PROGRAM prg_Piston
VAR
	fbPiston: FB_Piston;
	stPiston: ST_Piston;

	bPis_Next_P: BOOL;
	bPis_Next_N: BOOL;

	

	
	TON_0: TON;
	TON_1: TON;
	TON_2: TON;
	TON_3: TON;
	TON_4: TON;
	TON_5: TON;	
	i: INT;
END_VAR

act_InterLock();
act_Call_list_TanksMarinade();
act_Call_list_TanksColor();
act_Call_list_TanksCoolant();
act_Call_List_LineSource();
act_Call_List_LineTarget();
act_Call_list_CIP_SourceNTarget();
act_Call_list_CIP_Client();
act_Call_list_CIP_Tanks();
act_Call_list_Water();
act_Call_list_TriBlender_Selector();


IF bPis_Next_P THEN;
	m_Get_Next_P(iSel:=iPis_sel);
	bPis_Next_P:=FALSE;
END_IF

IF bPis_Next_N THEN;
	m_Get_Next_N(iSel:=iPis_sel);
	bPis_Next_N:=FALSE;
END_IF

FOR i:=0 TO E_Pis_Name.last DO
	ePisNameList:=i;
	arPisNameList[i]:=TO_STRING(ePisNameList);
END_FOR

ACTION act_Call_list_CIP_Client:
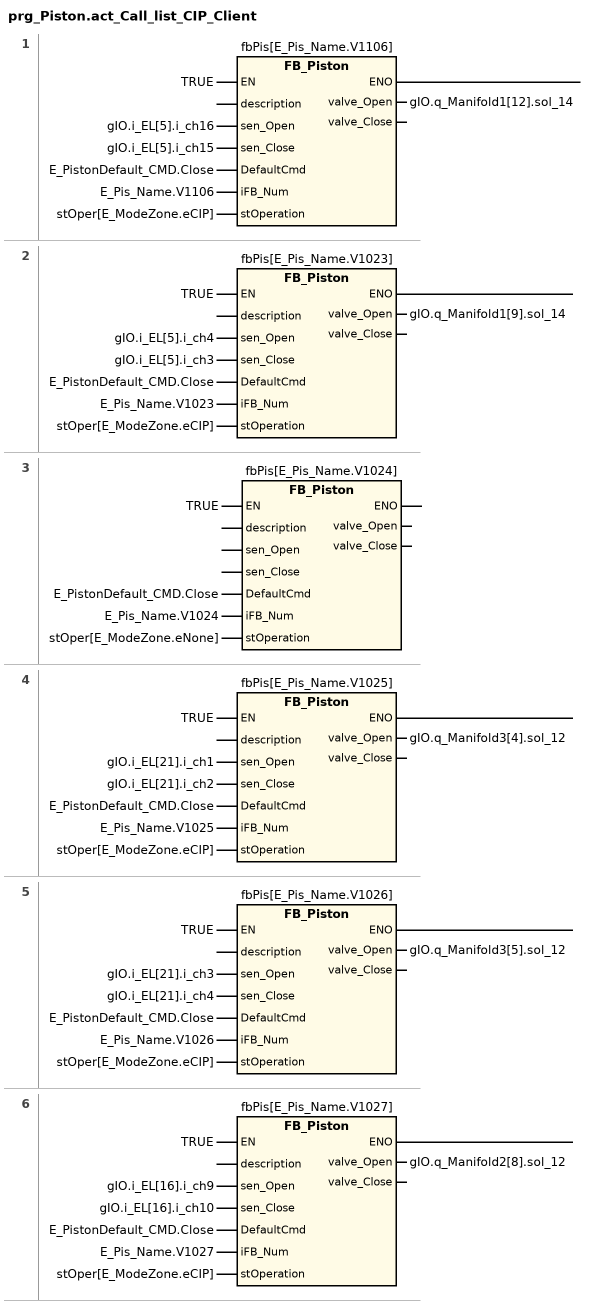
// NETWORK 1
fbPis[E_Pis_Name.V1106](
    sen_Open := gIO.i_EL[5].i_ch16,
    sen_Close := gIO.i_EL[5].i_ch15,
    DefaultCmd := E_PistonDefault_CMD.Close,
    iFB_Num := E_Pis_Name.V1106,
    stOperation := stOper[E_ModeZone.eCIP],
    valve_Open => gIO.q_Manifold1[12].sol_14); // FB_Piston

// NETWORK 2
fbPis[E_Pis_Name.V1023](
    sen_Open := gIO.i_EL[5].i_ch4,
    sen_Close := gIO.i_EL[5].i_ch3,
    DefaultCmd := E_PistonDefault_CMD.Close,
    iFB_Num := E_Pis_Name.V1023,
    stOperation := stOper[E_ModeZone.eCIP],
    valve_Open => gIO.q_Manifold1[9].sol_14); // FB_Piston

// NETWORK 3
fbPis[E_Pis_Name.V1024](
    DefaultCmd := E_PistonDefault_CMD.Close,
    iFB_Num := E_Pis_Name.V1024,
    stOperation := stOper[E_ModeZone.eNone]); // FB_Piston

// NETWORK 4
fbPis[E_Pis_Name.V1025](
    sen_Open := gIO.i_EL[21].i_ch1,
    sen_Close := gIO.i_EL[21].i_ch2,
    DefaultCmd := E_PistonDefault_CMD.Close,
    iFB_Num := E_Pis_Name.V1025,
    stOperation := stOper[E_ModeZone.eCIP],
    valve_Open => gIO.q_Manifold3[4].sol_12); // FB_Piston

// NETWORK 5
fbPis[E_Pis_Name.V1026](
    sen_Open := gIO.i_EL[21].i_ch3,
    sen_Close := gIO.i_EL[21].i_ch4,
    DefaultCmd := E_PistonDefault_CMD.Close,
    iFB_Num := E_Pis_Name.V1026,
    stOperation := stOper[E_ModeZone.eCIP],
    valve_Open => gIO.q_Manifold3[5].sol_12); // FB_Piston

// NETWORK 6
fbPis[E_Pis_Name.V1027](
    sen_Open := gIO.i_EL[16].i_ch9,
    sen_Close := gIO.i_EL[16].i_ch10,
    DefaultCmd := E_PistonDefault_CMD.Close,
    iFB_Num := E_Pis_Name.V1027,
    stOperation := stOper[E_ModeZone.eCIP],
    valve_Open => gIO.q_Manifold2[8].sol_12); // FB_Piston

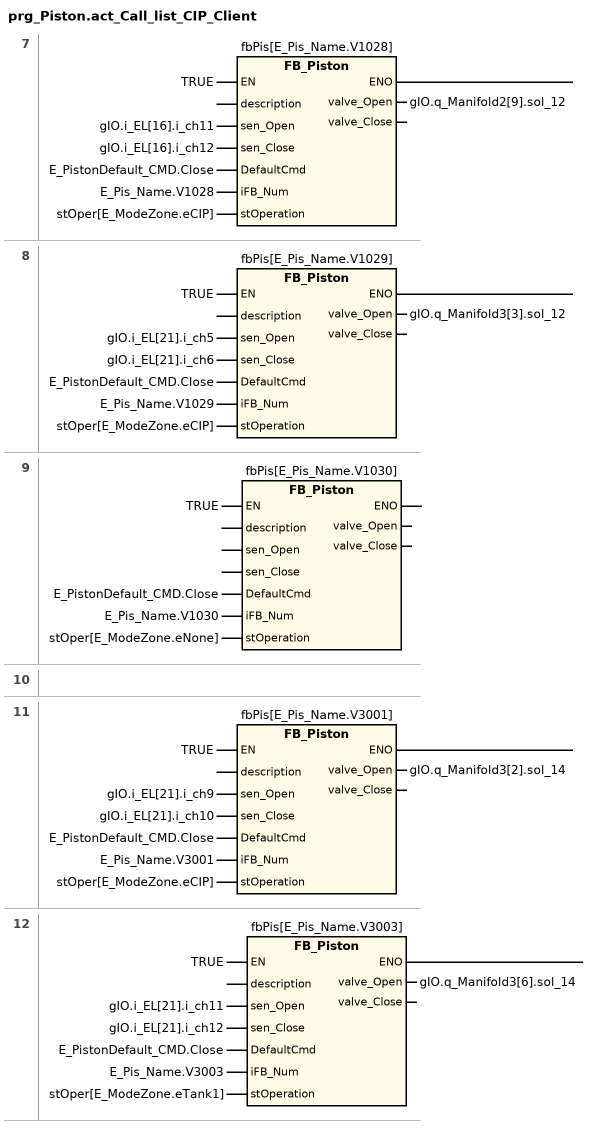
// NETWORK 7
fbPis[E_Pis_Name.V1028](
    sen_Open := gIO.i_EL[16].i_ch11,
    sen_Close := gIO.i_EL[16].i_ch12,
    DefaultCmd := E_PistonDefault_CMD.Close,
    iFB_Num := E_Pis_Name.V1028,
    stOperation := stOper[E_ModeZone.eCIP],
    valve_Open => gIO.q_Manifold2[9].sol_12); // FB_Piston

// NETWORK 8
fbPis[E_Pis_Name.V1029](
    sen_Open := gIO.i_EL[21].i_ch5,
    sen_Close := gIO.i_EL[21].i_ch6,
    DefaultCmd := E_PistonDefault_CMD.Close,
    iFB_Num := E_Pis_Name.V1029,
    stOperation := stOper[E_ModeZone.eCIP],
    valve_Open => gIO.q_Manifold3[3].sol_12); // FB_Piston

// NETWORK 9
fbPis[E_Pis_Name.V1030](
    DefaultCmd := E_PistonDefault_CMD.Close,
    iFB_Num := E_Pis_Name.V1030,
    stOperation := stOper[E_ModeZone.eNone]); // FB_Piston

// NETWORK 10

// NETWORK 11
fbPis[E_Pis_Name.V3001](
    sen_Open := gIO.i_EL[21].i_ch9,
    sen_Close := gIO.i_EL[21].i_ch10,
    DefaultCmd := E_PistonDefault_CMD.Close,
    iFB_Num := E_Pis_Name.V3001,
    stOperation := stOper[E_ModeZone.eCIP],
    valve_Open => gIO.q_Manifold3[2].sol_14); // FB_Piston

// NETWORK 12
fbPis[E_Pis_Name.V3003](
    sen_Open := gIO.i_EL[21].i_ch11,
    sen_Close := gIO.i_EL[21].i_ch12,
    DefaultCmd := E_PistonDefault_CMD.Close,
    iFB_Num := E_Pis_Name.V3003,
    stOperation := stOper[E_ModeZone.eTank1],
    valve_Open => gIO.q_Manifold3[6].sol_14); // FB_Piston

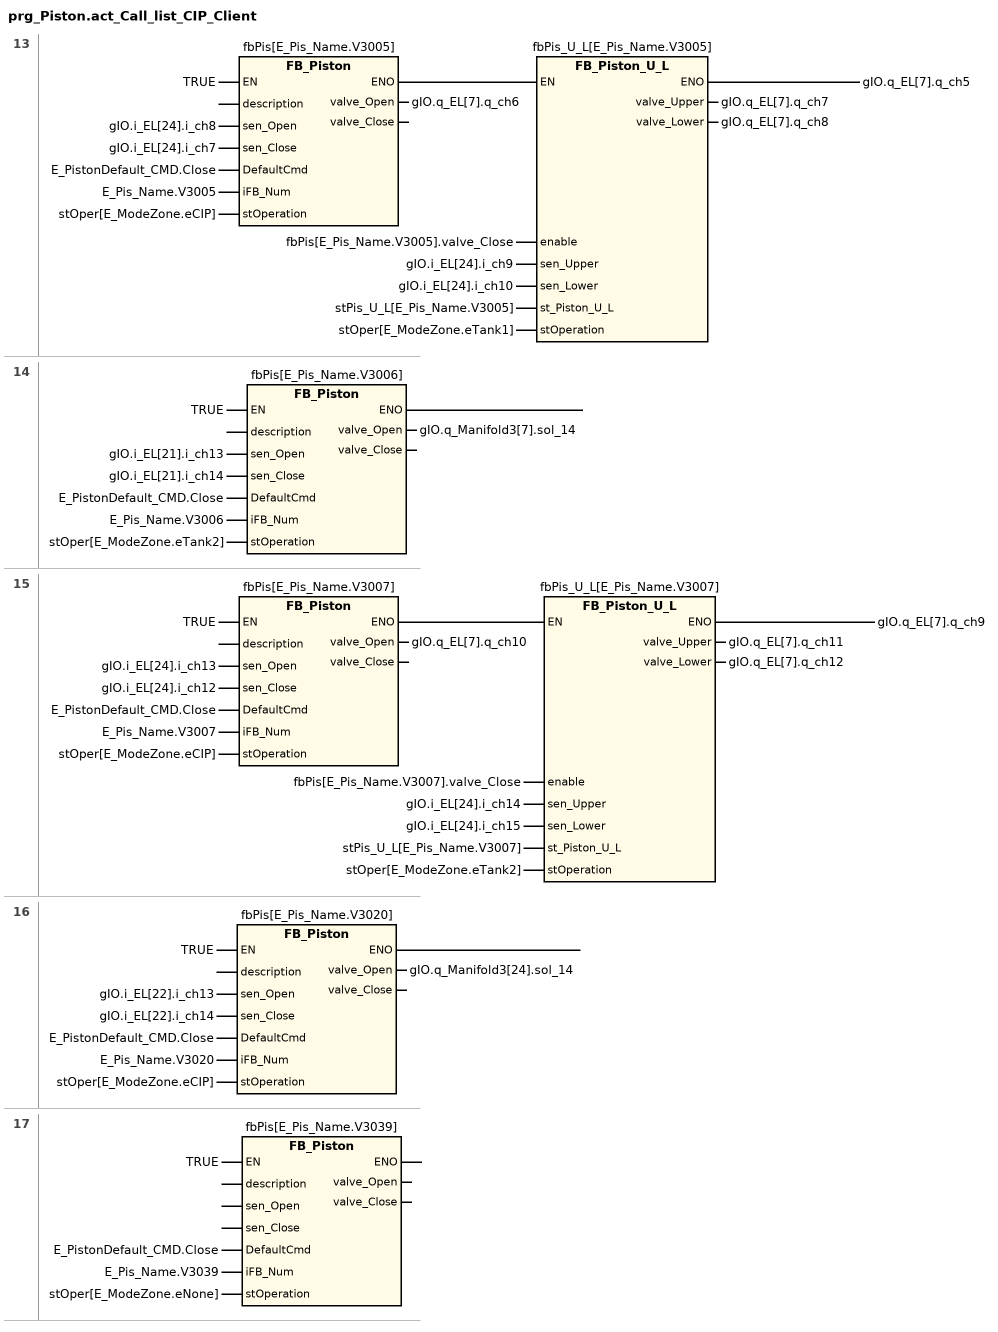
// NETWORK 13
fbPis[E_Pis_Name.V3005](
    sen_Open := gIO.i_EL[24].i_ch8,
    sen_Close := gIO.i_EL[24].i_ch7,
    DefaultCmd := E_PistonDefault_CMD.Close,
    iFB_Num := E_Pis_Name.V3005,
    stOperation := stOper[E_ModeZone.eCIP],
    valve_Open => gIO.q_EL[7].q_ch6); // FB_Piston
fbPis_U_L[E_Pis_Name.V3005](
    enable := fbPis[E_Pis_Name.V3005].valve_Close,
    sen_Upper := gIO.i_EL[24].i_ch9,
    sen_Lower := gIO.i_EL[24].i_ch10,
    st_Piston_U_L := stPis_U_L[E_Pis_Name.V3005],
    stOperation := stOper[E_ModeZone.eTank1],
    valve_Upper => gIO.q_EL[7].q_ch7,
    valve_Lower => gIO.q_EL[7].q_ch8); // FB_Piston_U_L
gIO.q_EL[7].q_ch5 := TRUE;

// NETWORK 14
fbPis[E_Pis_Name.V3006](
    sen_Open := gIO.i_EL[21].i_ch13,
    sen_Close := gIO.i_EL[21].i_ch14,
    DefaultCmd := E_PistonDefault_CMD.Close,
    iFB_Num := E_Pis_Name.V3006,
    stOperation := stOper[E_ModeZone.eTank2],
    valve_Open => gIO.q_Manifold3[7].sol_14); // FB_Piston

// NETWORK 15
fbPis[E_Pis_Name.V3007](
    sen_Open := gIO.i_EL[24].i_ch13,
    sen_Close := gIO.i_EL[24].i_ch12,
    DefaultCmd := E_PistonDefault_CMD.Close,
    iFB_Num := E_Pis_Name.V3007,
    stOperation := stOper[E_ModeZone.eCIP],
    valve_Open => gIO.q_EL[7].q_ch10); // FB_Piston
fbPis_U_L[E_Pis_Name.V3007](
    enable := fbPis[E_Pis_Name.V3007].valve_Close,
    sen_Upper := gIO.i_EL[24].i_ch14,
    sen_Lower := gIO.i_EL[24].i_ch15,
    st_Piston_U_L := stPis_U_L[E_Pis_Name.V3007],
    stOperation := stOper[E_ModeZone.eTank2],
    valve_Upper => gIO.q_EL[7].q_ch11,
    valve_Lower => gIO.q_EL[7].q_ch12); // FB_Piston_U_L
gIO.q_EL[7].q_ch9 := TRUE;

// NETWORK 16
fbPis[E_Pis_Name.V3020](
    sen_Open := gIO.i_EL[22].i_ch13,
    sen_Close := gIO.i_EL[22].i_ch14,
    DefaultCmd := E_PistonDefault_CMD.Close,
    iFB_Num := E_Pis_Name.V3020,
    stOperation := stOper[E_ModeZone.eCIP],
    valve_Open => gIO.q_Manifold3[24].sol_14); // FB_Piston

// NETWORK 17
fbPis[E_Pis_Name.V3039](
    DefaultCmd := E_PistonDefault_CMD.Close,
    iFB_Num := E_Pis_Name.V3039,
    stOperation := stOper[E_ModeZone.eNone]); // FB_Piston

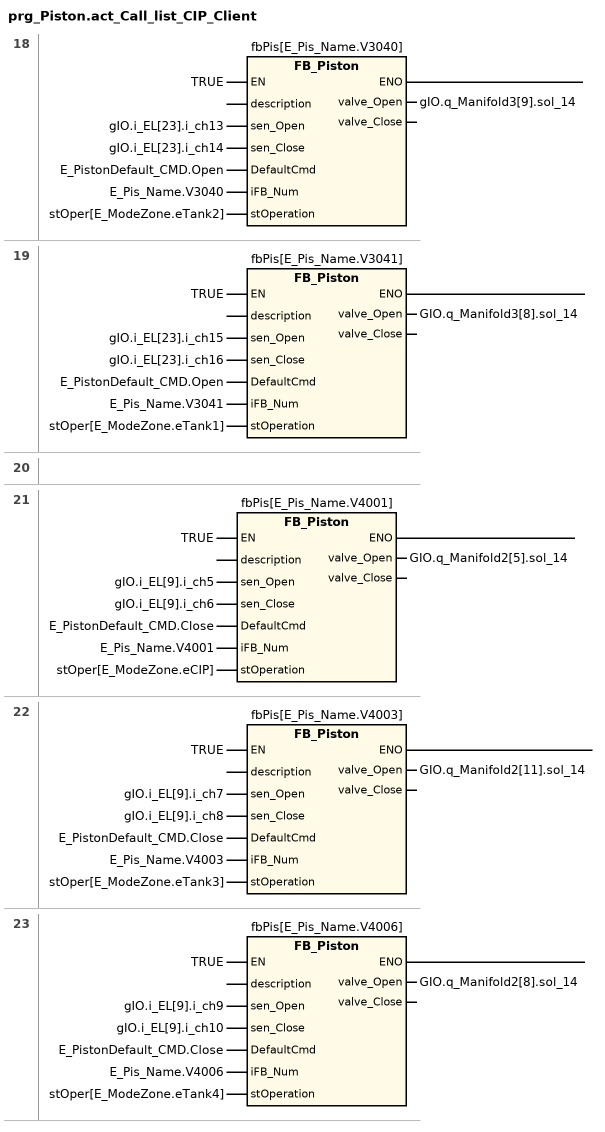
// NETWORK 18
fbPis[E_Pis_Name.V3040](
    sen_Open := gIO.i_EL[23].i_ch13,
    sen_Close := gIO.i_EL[23].i_ch14,
    DefaultCmd := E_PistonDefault_CMD.Open,
    iFB_Num := E_Pis_Name.V3040,
    stOperation := stOper[E_ModeZone.eTank2],
    valve_Open => gIO.q_Manifold3[9].sol_14); // FB_Piston

// NETWORK 19
fbPis[E_Pis_Name.V3041](
    sen_Open := gIO.i_EL[23].i_ch15,
    sen_Close := gIO.i_EL[23].i_ch16,
    DefaultCmd := E_PistonDefault_CMD.Open,
    iFB_Num := E_Pis_Name.V3041,
    stOperation := stOper[E_ModeZone.eTank1],
    valve_Open => GIO.q_Manifold3[8].sol_14); // FB_Piston

// NETWORK 20

// NETWORK 21
fbPis[E_Pis_Name.V4001](
    sen_Open := gIO.i_EL[9].i_ch5,
    sen_Close := gIO.i_EL[9].i_ch6,
    DefaultCmd := E_PistonDefault_CMD.Close,
    iFB_Num := E_Pis_Name.V4001,
    stOperation := stOper[E_ModeZone.eCIP],
    valve_Open => GIO.q_Manifold2[5].sol_14); // FB_Piston

// NETWORK 22
fbPis[E_Pis_Name.V4003](
    sen_Open := gIO.i_EL[9].i_ch7,
    sen_Close := gIO.i_EL[9].i_ch8,
    DefaultCmd := E_PistonDefault_CMD.Close,
    iFB_Num := E_Pis_Name.V4003,
    stOperation := stOper[E_ModeZone.eTank3],
    valve_Open => GIO.q_Manifold2[11].sol_14); // FB_Piston

// NETWORK 23
fbPis[E_Pis_Name.V4006](
    sen_Open := gIO.i_EL[9].i_ch9,
    sen_Close := gIO.i_EL[9].i_ch10,
    DefaultCmd := E_PistonDefault_CMD.Close,
    iFB_Num := E_Pis_Name.V4006,
    stOperation := stOper[E_ModeZone.eTank4],
    valve_Open => GIO.q_Manifold2[8].sol_14); // FB_Piston

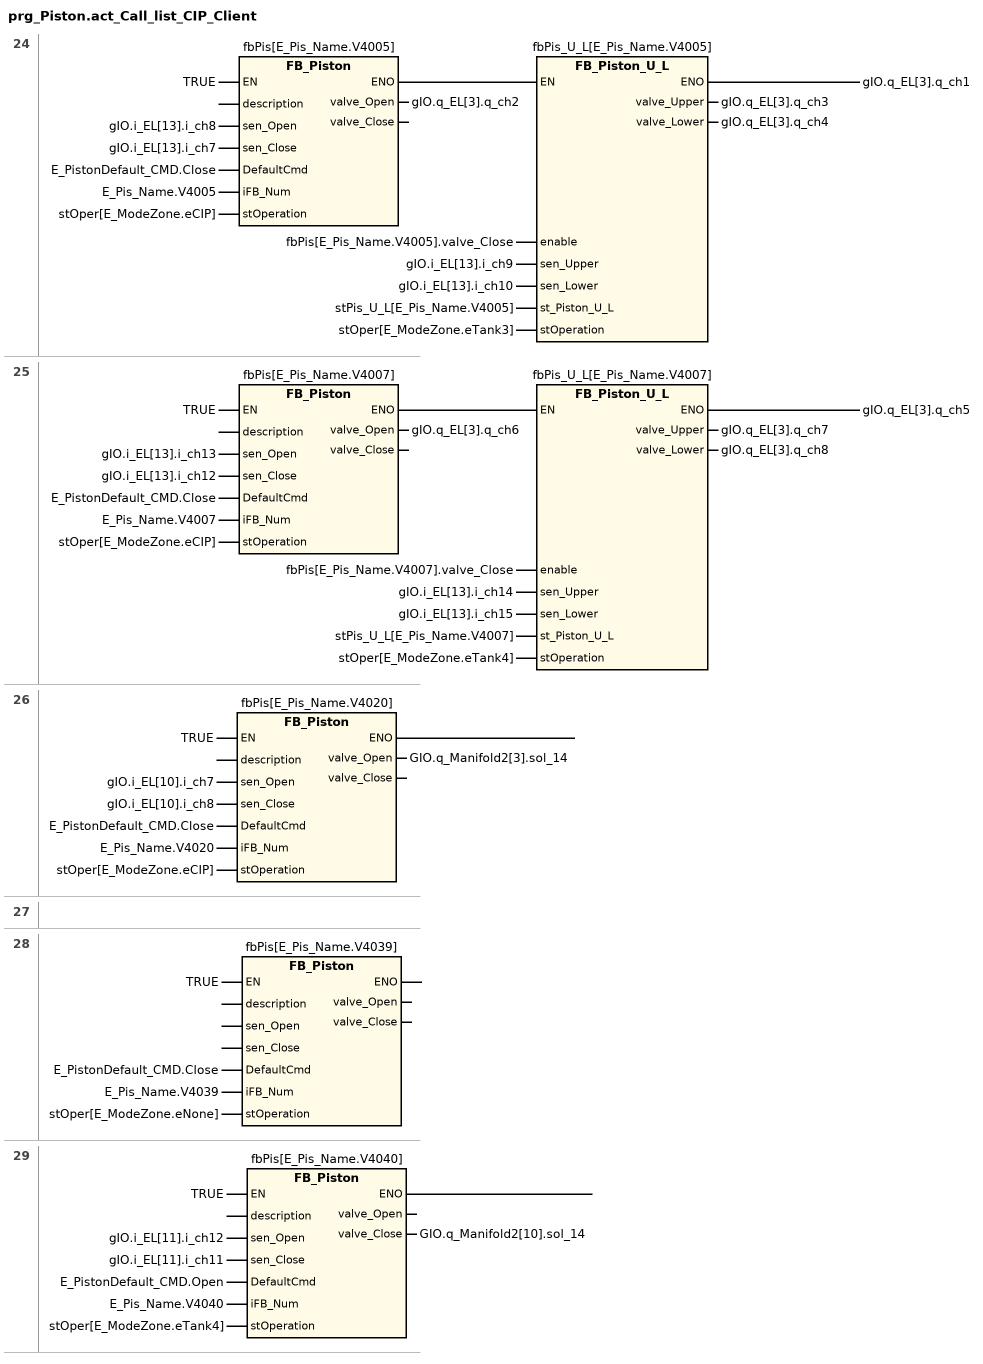
// NETWORK 24
fbPis[E_Pis_Name.V4005](
    sen_Open := gIO.i_EL[13].i_ch8,
    sen_Close := gIO.i_EL[13].i_ch7,
    DefaultCmd := E_PistonDefault_CMD.Close,
    iFB_Num := E_Pis_Name.V4005,
    stOperation := stOper[E_ModeZone.eCIP],
    valve_Open => gIO.q_EL[3].q_ch2); // FB_Piston
fbPis_U_L[E_Pis_Name.V4005](
    enable := fbPis[E_Pis_Name.V4005].valve_Close,
    sen_Upper := gIO.i_EL[13].i_ch9,
    sen_Lower := gIO.i_EL[13].i_ch10,
    st_Piston_U_L := stPis_U_L[E_Pis_Name.V4005],
    stOperation := stOper[E_ModeZone.eTank3],
    valve_Upper => gIO.q_EL[3].q_ch3,
    valve_Lower => gIO.q_EL[3].q_ch4); // FB_Piston_U_L
gIO.q_EL[3].q_ch1 := TRUE;

// NETWORK 25
fbPis[E_Pis_Name.V4007](
    sen_Open := gIO.i_EL[13].i_ch13,
    sen_Close := gIO.i_EL[13].i_ch12,
    DefaultCmd := E_PistonDefault_CMD.Close,
    iFB_Num := E_Pis_Name.V4007,
    stOperation := stOper[E_ModeZone.eCIP],
    valve_Open => gIO.q_EL[3].q_ch6); // FB_Piston
fbPis_U_L[E_Pis_Name.V4007](
    enable := fbPis[E_Pis_Name.V4007].valve_Close,
    sen_Upper := gIO.i_EL[13].i_ch14,
    sen_Lower := gIO.i_EL[13].i_ch15,
    st_Piston_U_L := stPis_U_L[E_Pis_Name.V4007],
    stOperation := stOper[E_ModeZone.eTank4],
    valve_Upper => gIO.q_EL[3].q_ch7,
    valve_Lower => gIO.q_EL[3].q_ch8); // FB_Piston_U_L
gIO.q_EL[3].q_ch5 := TRUE;

// NETWORK 26
fbPis[E_Pis_Name.V4020](
    sen_Open := gIO.i_EL[10].i_ch7,
    sen_Close := gIO.i_EL[10].i_ch8,
    DefaultCmd := E_PistonDefault_CMD.Close,
    iFB_Num := E_Pis_Name.V4020,
    stOperation := stOper[E_ModeZone.eCIP],
    valve_Open => GIO.q_Manifold2[3].sol_14); // FB_Piston

// NETWORK 27

// NETWORK 28
fbPis[E_Pis_Name.V4039](
    DefaultCmd := E_PistonDefault_CMD.Close,
    iFB_Num := E_Pis_Name.V4039,
    stOperation := stOper[E_ModeZone.eNone]); // FB_Piston

// NETWORK 29
fbPis[E_Pis_Name.V4040](
    sen_Open := gIO.i_EL[11].i_ch12,
    sen_Close := gIO.i_EL[11].i_ch11,
    DefaultCmd := E_PistonDefault_CMD.Open,
    iFB_Num := E_Pis_Name.V4040,
    stOperation := stOper[E_ModeZone.eTank4],
    valve_Close => GIO.q_Manifold2[10].sol_14); // FB_Piston

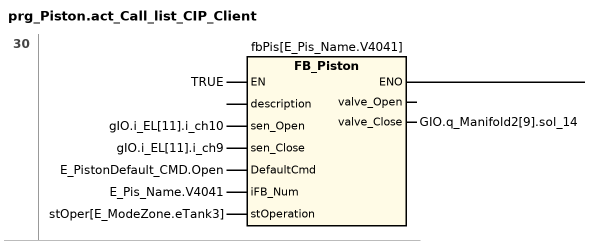
// NETWORK 30
fbPis[E_Pis_Name.V4041](
    sen_Open := gIO.i_EL[11].i_ch10,
    sen_Close := gIO.i_EL[11].i_ch9,
    DefaultCmd := E_PistonDefault_CMD.Open,
    iFB_Num := E_Pis_Name.V4041,
    stOperation := stOper[E_ModeZone.eTank3],
    valve_Close => GIO.q_Manifold2[9].sol_14); // FB_Piston
END_ACTION

ACTION act_Call_list_CIP_SourceNTarget:
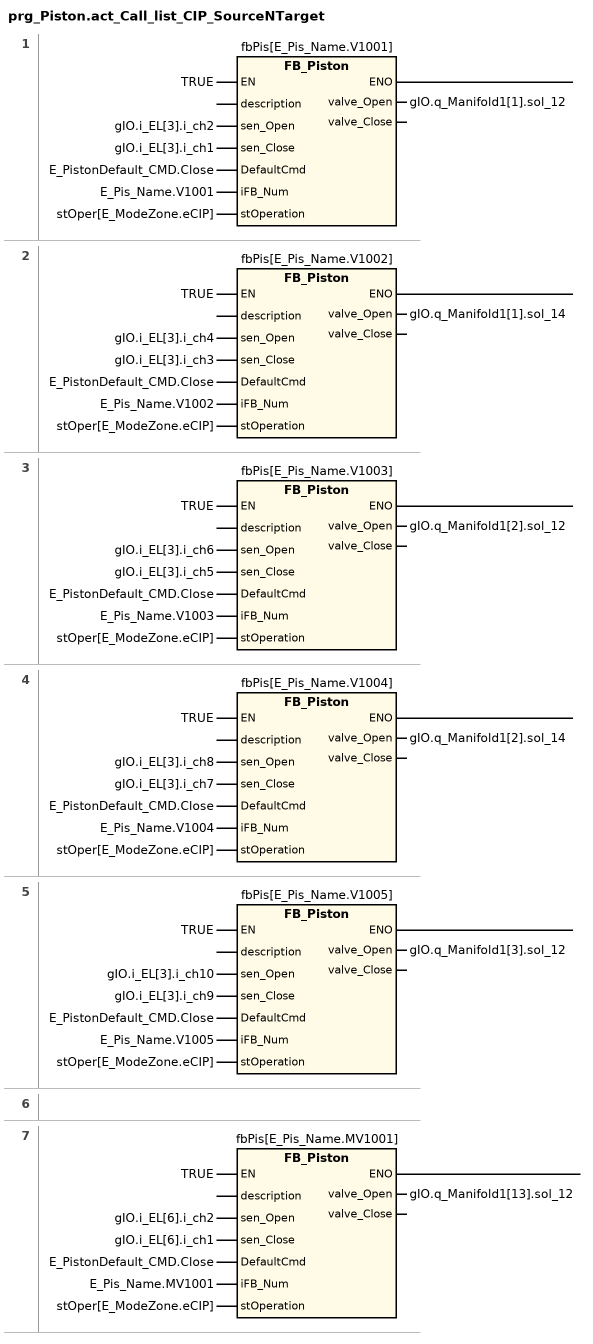
// NETWORK 1
fbPis[E_Pis_Name.V1001](
    sen_Open := gIO.i_EL[3].i_ch2,
    sen_Close := gIO.i_EL[3].i_ch1,
    DefaultCmd := E_PistonDefault_CMD.Close,
    iFB_Num := E_Pis_Name.V1001,
    stOperation := stOper[E_ModeZone.eCIP],
    valve_Open => gIO.q_Manifold1[1].sol_12); // FB_Piston

// NETWORK 2
fbPis[E_Pis_Name.V1002](
    sen_Open := gIO.i_EL[3].i_ch4,
    sen_Close := gIO.i_EL[3].i_ch3,
    DefaultCmd := E_PistonDefault_CMD.Close,
    iFB_Num := E_Pis_Name.V1002,
    stOperation := stOper[E_ModeZone.eCIP],
    valve_Open => gIO.q_Manifold1[1].sol_14); // FB_Piston

// NETWORK 3
fbPis[E_Pis_Name.V1003](
    sen_Open := gIO.i_EL[3].i_ch6,
    sen_Close := gIO.i_EL[3].i_ch5,
    DefaultCmd := E_PistonDefault_CMD.Close,
    iFB_Num := E_Pis_Name.V1003,
    stOperation := stOper[E_ModeZone.eCIP],
    valve_Open => gIO.q_Manifold1[2].sol_12); // FB_Piston

// NETWORK 4
fbPis[E_Pis_Name.V1004](
    sen_Open := gIO.i_EL[3].i_ch8,
    sen_Close := gIO.i_EL[3].i_ch7,
    DefaultCmd := E_PistonDefault_CMD.Close,
    iFB_Num := E_Pis_Name.V1004,
    stOperation := stOper[E_ModeZone.eCIP],
    valve_Open => gIO.q_Manifold1[2].sol_14); // FB_Piston

// NETWORK 5
fbPis[E_Pis_Name.V1005](
    sen_Open := gIO.i_EL[3].i_ch10,
    sen_Close := gIO.i_EL[3].i_ch9,
    DefaultCmd := E_PistonDefault_CMD.Close,
    iFB_Num := E_Pis_Name.V1005,
    stOperation := stOper[E_ModeZone.eCIP],
    valve_Open => gIO.q_Manifold1[3].sol_12); // FB_Piston

// NETWORK 6

// NETWORK 7
fbPis[E_Pis_Name.MV1001](
    sen_Open := gIO.i_EL[6].i_ch2,
    sen_Close := gIO.i_EL[6].i_ch1,
    DefaultCmd := E_PistonDefault_CMD.Close,
    iFB_Num := E_Pis_Name.MV1001,
    stOperation := stOper[E_ModeZone.eCIP],
    valve_Open => gIO.q_Manifold1[13].sol_12); // FB_Piston

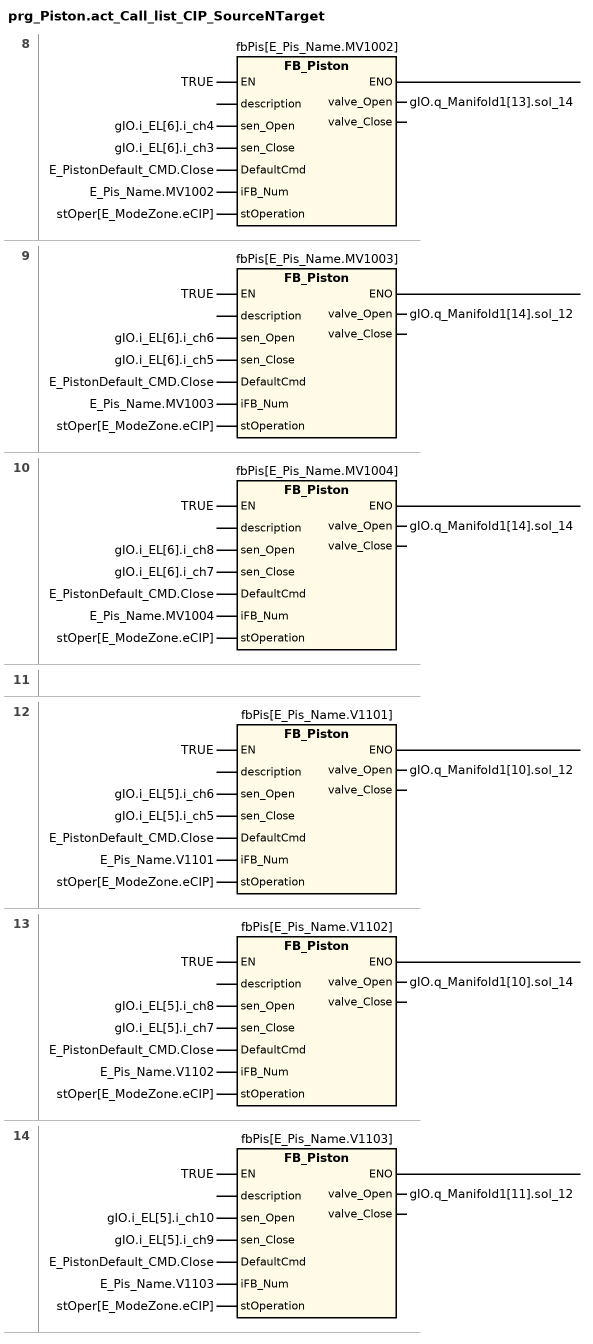
// NETWORK 8
fbPis[E_Pis_Name.MV1002](
    sen_Open := gIO.i_EL[6].i_ch4,
    sen_Close := gIO.i_EL[6].i_ch3,
    DefaultCmd := E_PistonDefault_CMD.Close,
    iFB_Num := E_Pis_Name.MV1002,
    stOperation := stOper[E_ModeZone.eCIP],
    valve_Open => gIO.q_Manifold1[13].sol_14); // FB_Piston

// NETWORK 9
fbPis[E_Pis_Name.MV1003](
    sen_Open := gIO.i_EL[6].i_ch6,
    sen_Close := gIO.i_EL[6].i_ch5,
    DefaultCmd := E_PistonDefault_CMD.Close,
    iFB_Num := E_Pis_Name.MV1003,
    stOperation := stOper[E_ModeZone.eCIP],
    valve_Open => gIO.q_Manifold1[14].sol_12); // FB_Piston

// NETWORK 10
fbPis[E_Pis_Name.MV1004](
    sen_Open := gIO.i_EL[6].i_ch8,
    sen_Close := gIO.i_EL[6].i_ch7,
    DefaultCmd := E_PistonDefault_CMD.Close,
    iFB_Num := E_Pis_Name.MV1004,
    stOperation := stOper[E_ModeZone.eCIP],
    valve_Open => gIO.q_Manifold1[14].sol_14); // FB_Piston

// NETWORK 11

// NETWORK 12
fbPis[E_Pis_Name.V1101](
    sen_Open := gIO.i_EL[5].i_ch6,
    sen_Close := gIO.i_EL[5].i_ch5,
    DefaultCmd := E_PistonDefault_CMD.Close,
    iFB_Num := E_Pis_Name.V1101,
    stOperation := stOper[E_ModeZone.eCIP],
    valve_Open => gIO.q_Manifold1[10].sol_12); // FB_Piston

// NETWORK 13
fbPis[E_Pis_Name.V1102](
    sen_Open := gIO.i_EL[5].i_ch8,
    sen_Close := gIO.i_EL[5].i_ch7,
    DefaultCmd := E_PistonDefault_CMD.Close,
    iFB_Num := E_Pis_Name.V1102,
    stOperation := stOper[E_ModeZone.eCIP],
    valve_Open => gIO.q_Manifold1[10].sol_14); // FB_Piston

// NETWORK 14
fbPis[E_Pis_Name.V1103](
    sen_Open := gIO.i_EL[5].i_ch10,
    sen_Close := gIO.i_EL[5].i_ch9,
    DefaultCmd := E_PistonDefault_CMD.Close,
    iFB_Num := E_Pis_Name.V1103,
    stOperation := stOper[E_ModeZone.eCIP],
    valve_Open => gIO.q_Manifold1[11].sol_12); // FB_Piston

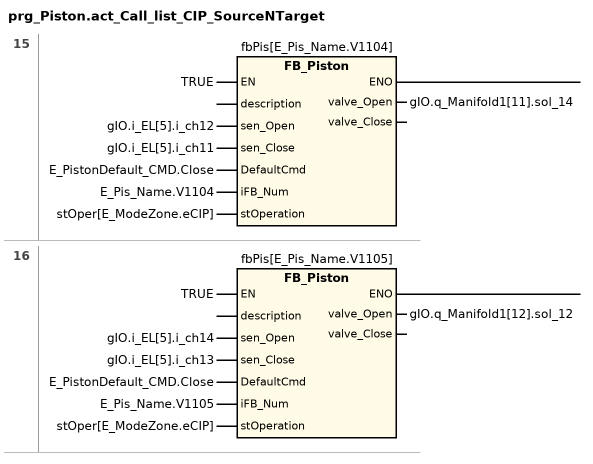
// NETWORK 15
fbPis[E_Pis_Name.V1104](
    sen_Open := gIO.i_EL[5].i_ch12,
    sen_Close := gIO.i_EL[5].i_ch11,
    DefaultCmd := E_PistonDefault_CMD.Close,
    iFB_Num := E_Pis_Name.V1104,
    stOperation := stOper[E_ModeZone.eCIP],
    valve_Open => gIO.q_Manifold1[11].sol_14); // FB_Piston

// NETWORK 16
fbPis[E_Pis_Name.V1105](
    sen_Open := gIO.i_EL[5].i_ch14,
    sen_Close := gIO.i_EL[5].i_ch13,
    DefaultCmd := E_PistonDefault_CMD.Close,
    iFB_Num := E_Pis_Name.V1105,
    stOperation := stOper[E_ModeZone.eCIP],
    valve_Open => gIO.q_Manifold1[12].sol_12); // FB_Piston
END_ACTION

ACTION act_Call_list_CIP_Tanks:
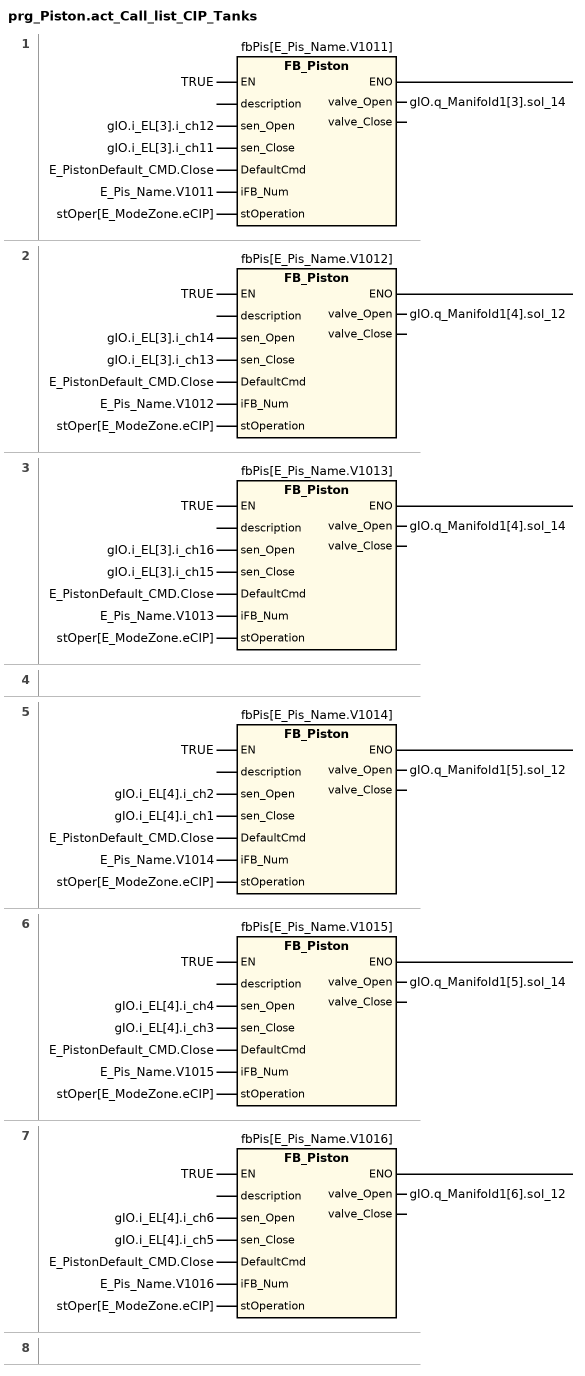
// NETWORK 1
fbPis[E_Pis_Name.V1011](
    sen_Open := gIO.i_EL[3].i_ch12,
    sen_Close := gIO.i_EL[3].i_ch11,
    DefaultCmd := E_PistonDefault_CMD.Close,
    iFB_Num := E_Pis_Name.V1011,
    stOperation := stOper[E_ModeZone.eCIP],
    valve_Open => gIO.q_Manifold1[3].sol_14); // FB_Piston

// NETWORK 2
fbPis[E_Pis_Name.V1012](
    sen_Open := gIO.i_EL[3].i_ch14,
    sen_Close := gIO.i_EL[3].i_ch13,
    DefaultCmd := E_PistonDefault_CMD.Close,
    iFB_Num := E_Pis_Name.V1012,
    stOperation := stOper[E_ModeZone.eCIP],
    valve_Open => gIO.q_Manifold1[4].sol_12); // FB_Piston

// NETWORK 3
fbPis[E_Pis_Name.V1013](
    sen_Open := gIO.i_EL[3].i_ch16,
    sen_Close := gIO.i_EL[3].i_ch15,
    DefaultCmd := E_PistonDefault_CMD.Close,
    iFB_Num := E_Pis_Name.V1013,
    stOperation := stOper[E_ModeZone.eCIP],
    valve_Open => gIO.q_Manifold1[4].sol_14); // FB_Piston

// NETWORK 4

// NETWORK 5
fbPis[E_Pis_Name.V1014](
    sen_Open := gIO.i_EL[4].i_ch2,
    sen_Close := gIO.i_EL[4].i_ch1,
    DefaultCmd := E_PistonDefault_CMD.Close,
    iFB_Num := E_Pis_Name.V1014,
    stOperation := stOper[E_ModeZone.eCIP],
    valve_Open => gIO.q_Manifold1[5].sol_12); // FB_Piston

// NETWORK 6
fbPis[E_Pis_Name.V1015](
    sen_Open := gIO.i_EL[4].i_ch4,
    sen_Close := gIO.i_EL[4].i_ch3,
    DefaultCmd := E_PistonDefault_CMD.Close,
    iFB_Num := E_Pis_Name.V1015,
    stOperation := stOper[E_ModeZone.eCIP],
    valve_Open => gIO.q_Manifold1[5].sol_14); // FB_Piston

// NETWORK 7
fbPis[E_Pis_Name.V1016](
    sen_Open := gIO.i_EL[4].i_ch6,
    sen_Close := gIO.i_EL[4].i_ch5,
    DefaultCmd := E_PistonDefault_CMD.Close,
    iFB_Num := E_Pis_Name.V1016,
    stOperation := stOper[E_ModeZone.eCIP],
    valve_Open => gIO.q_Manifold1[6].sol_12); // FB_Piston

// NETWORK 8

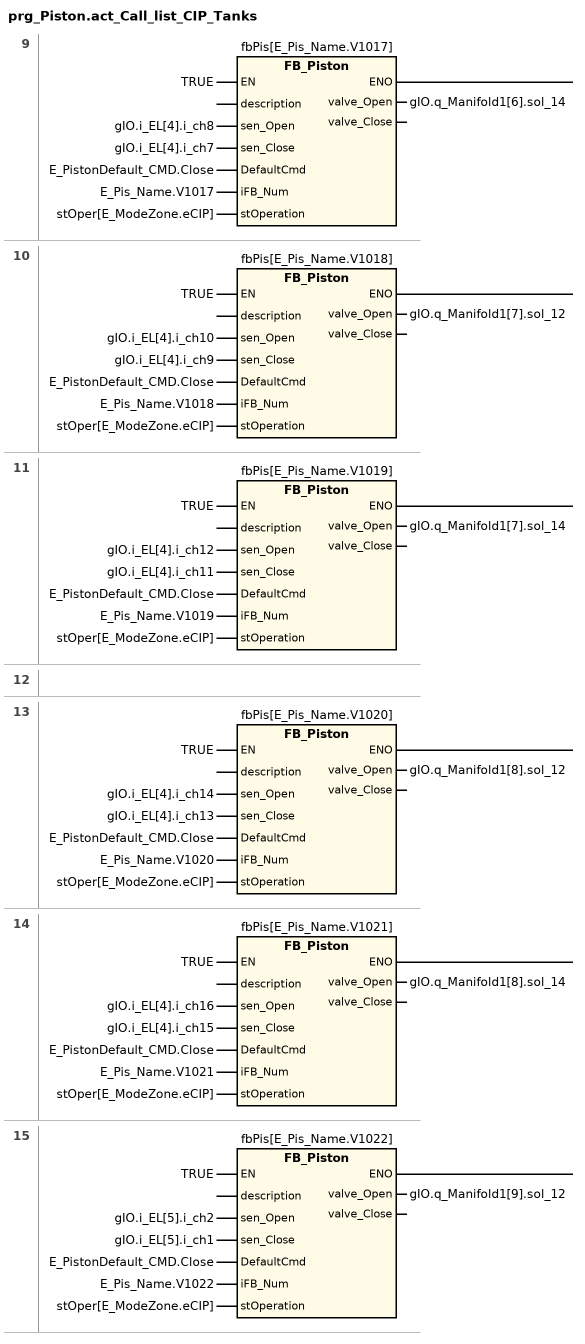
// NETWORK 9
fbPis[E_Pis_Name.V1017](
    sen_Open := gIO.i_EL[4].i_ch8,
    sen_Close := gIO.i_EL[4].i_ch7,
    DefaultCmd := E_PistonDefault_CMD.Close,
    iFB_Num := E_Pis_Name.V1017,
    stOperation := stOper[E_ModeZone.eCIP],
    valve_Open => gIO.q_Manifold1[6].sol_14); // FB_Piston

// NETWORK 10
fbPis[E_Pis_Name.V1018](
    sen_Open := gIO.i_EL[4].i_ch10,
    sen_Close := gIO.i_EL[4].i_ch9,
    DefaultCmd := E_PistonDefault_CMD.Close,
    iFB_Num := E_Pis_Name.V1018,
    stOperation := stOper[E_ModeZone.eCIP],
    valve_Open => gIO.q_Manifold1[7].sol_12); // FB_Piston

// NETWORK 11
fbPis[E_Pis_Name.V1019](
    sen_Open := gIO.i_EL[4].i_ch12,
    sen_Close := gIO.i_EL[4].i_ch11,
    DefaultCmd := E_PistonDefault_CMD.Close,
    iFB_Num := E_Pis_Name.V1019,
    stOperation := stOper[E_ModeZone.eCIP],
    valve_Open => gIO.q_Manifold1[7].sol_14); // FB_Piston

// NETWORK 12

// NETWORK 13
fbPis[E_Pis_Name.V1020](
    sen_Open := gIO.i_EL[4].i_ch14,
    sen_Close := gIO.i_EL[4].i_ch13,
    DefaultCmd := E_PistonDefault_CMD.Close,
    iFB_Num := E_Pis_Name.V1020,
    stOperation := stOper[E_ModeZone.eCIP],
    valve_Open => gIO.q_Manifold1[8].sol_12); // FB_Piston

// NETWORK 14
fbPis[E_Pis_Name.V1021](
    sen_Open := gIO.i_EL[4].i_ch16,
    sen_Close := gIO.i_EL[4].i_ch15,
    DefaultCmd := E_PistonDefault_CMD.Close,
    iFB_Num := E_Pis_Name.V1021,
    stOperation := stOper[E_ModeZone.eCIP],
    valve_Open => gIO.q_Manifold1[8].sol_14); // FB_Piston

// NETWORK 15
fbPis[E_Pis_Name.V1022](
    sen_Open := gIO.i_EL[5].i_ch2,
    sen_Close := gIO.i_EL[5].i_ch1,
    DefaultCmd := E_PistonDefault_CMD.Close,
    iFB_Num := E_Pis_Name.V1022,
    stOperation := stOper[E_ModeZone.eCIP],
    valve_Open => gIO.q_Manifold1[9].sol_12); // FB_Piston

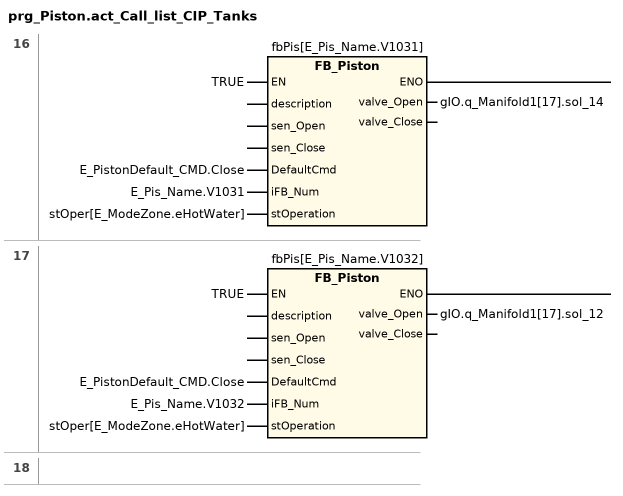
// NETWORK 16
fbPis[E_Pis_Name.V1031](
    DefaultCmd := E_PistonDefault_CMD.Close,
    iFB_Num := E_Pis_Name.V1031,
    stOperation := stOper[E_ModeZone.eHotWater],
    valve_Open => gIO.q_Manifold1[17].sol_14); // FB_Piston

// NETWORK 17
fbPis[E_Pis_Name.V1032](
    DefaultCmd := E_PistonDefault_CMD.Close,
    iFB_Num := E_Pis_Name.V1032,
    stOperation := stOper[E_ModeZone.eHotWater],
    valve_Open => gIO.q_Manifold1[17].sol_12); // FB_Piston

// NETWORK 18
END_ACTION

ACTION act_Call_List_LineSource:
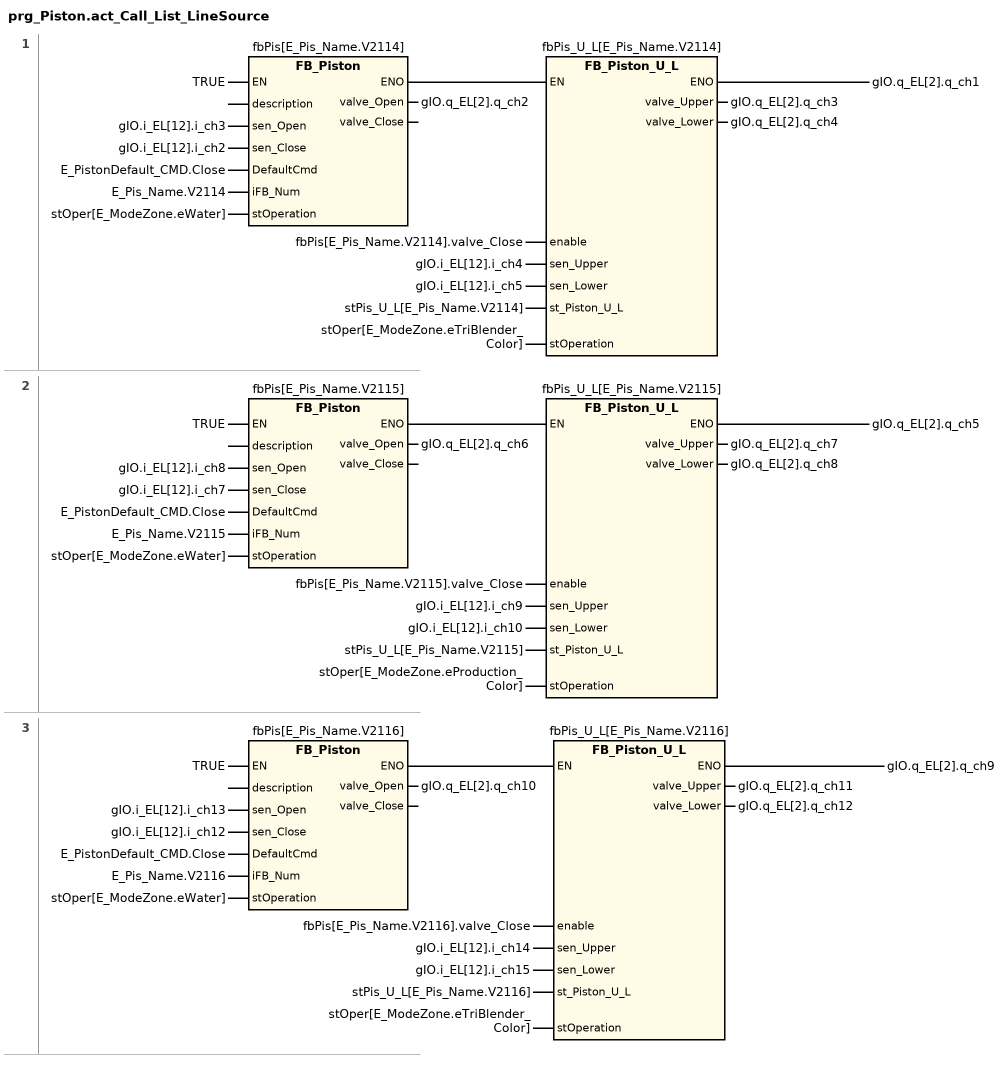
// NETWORK 1
fbPis[E_Pis_Name.V2114](
    sen_Open := gIO.i_EL[12].i_ch3,
    sen_Close := gIO.i_EL[12].i_ch2,
    DefaultCmd := E_PistonDefault_CMD.Close,
    iFB_Num := E_Pis_Name.V2114,
    stOperation := stOper[E_ModeZone.eWater],
    valve_Open => gIO.q_EL[2].q_ch2); // FB_Piston
fbPis_U_L[E_Pis_Name.V2114](
    enable := fbPis[E_Pis_Name.V2114].valve_Close,
    sen_Upper := gIO.i_EL[12].i_ch4,
    sen_Lower := gIO.i_EL[12].i_ch5,
    st_Piston_U_L := stPis_U_L[E_Pis_Name.V2114],
    stOperation := stOper[E_ModeZone.eTriBlender_Color],
    valve_Upper => gIO.q_EL[2].q_ch3,
    valve_Lower => gIO.q_EL[2].q_ch4); // FB_Piston_U_L
gIO.q_EL[2].q_ch1 := TRUE;

// NETWORK 2
fbPis[E_Pis_Name.V2115](
    sen_Open := gIO.i_EL[12].i_ch8,
    sen_Close := gIO.i_EL[12].i_ch7,
    DefaultCmd := E_PistonDefault_CMD.Close,
    iFB_Num := E_Pis_Name.V2115,
    stOperation := stOper[E_ModeZone.eWater],
    valve_Open => gIO.q_EL[2].q_ch6); // FB_Piston
fbPis_U_L[E_Pis_Name.V2115](
    enable := fbPis[E_Pis_Name.V2115].valve_Close,
    sen_Upper := gIO.i_EL[12].i_ch9,
    sen_Lower := gIO.i_EL[12].i_ch10,
    st_Piston_U_L := stPis_U_L[E_Pis_Name.V2115],
    stOperation := stOper[E_ModeZone.eProduction_Color],
    valve_Upper => gIO.q_EL[2].q_ch7,
    valve_Lower => gIO.q_EL[2].q_ch8); // FB_Piston_U_L
gIO.q_EL[2].q_ch5 := TRUE;

// NETWORK 3
fbPis[E_Pis_Name.V2116](
    sen_Open := gIO.i_EL[12].i_ch13,
    sen_Close := gIO.i_EL[12].i_ch12,
    DefaultCmd := E_PistonDefault_CMD.Close,
    iFB_Num := E_Pis_Name.V2116,
    stOperation := stOper[E_ModeZone.eWater],
    valve_Open => gIO.q_EL[2].q_ch10); // FB_Piston
fbPis_U_L[E_Pis_Name.V2116](
    enable := fbPis[E_Pis_Name.V2116].valve_Close,
    sen_Upper := gIO.i_EL[12].i_ch14,
    sen_Lower := gIO.i_EL[12].i_ch15,
    st_Piston_U_L := stPis_U_L[E_Pis_Name.V2116],
    stOperation := stOper[E_ModeZone.eTriBlender_Color],
    valve_Upper => gIO.q_EL[2].q_ch11,
    valve_Lower => gIO.q_EL[2].q_ch12); // FB_Piston_U_L
gIO.q_EL[2].q_ch9 := TRUE;

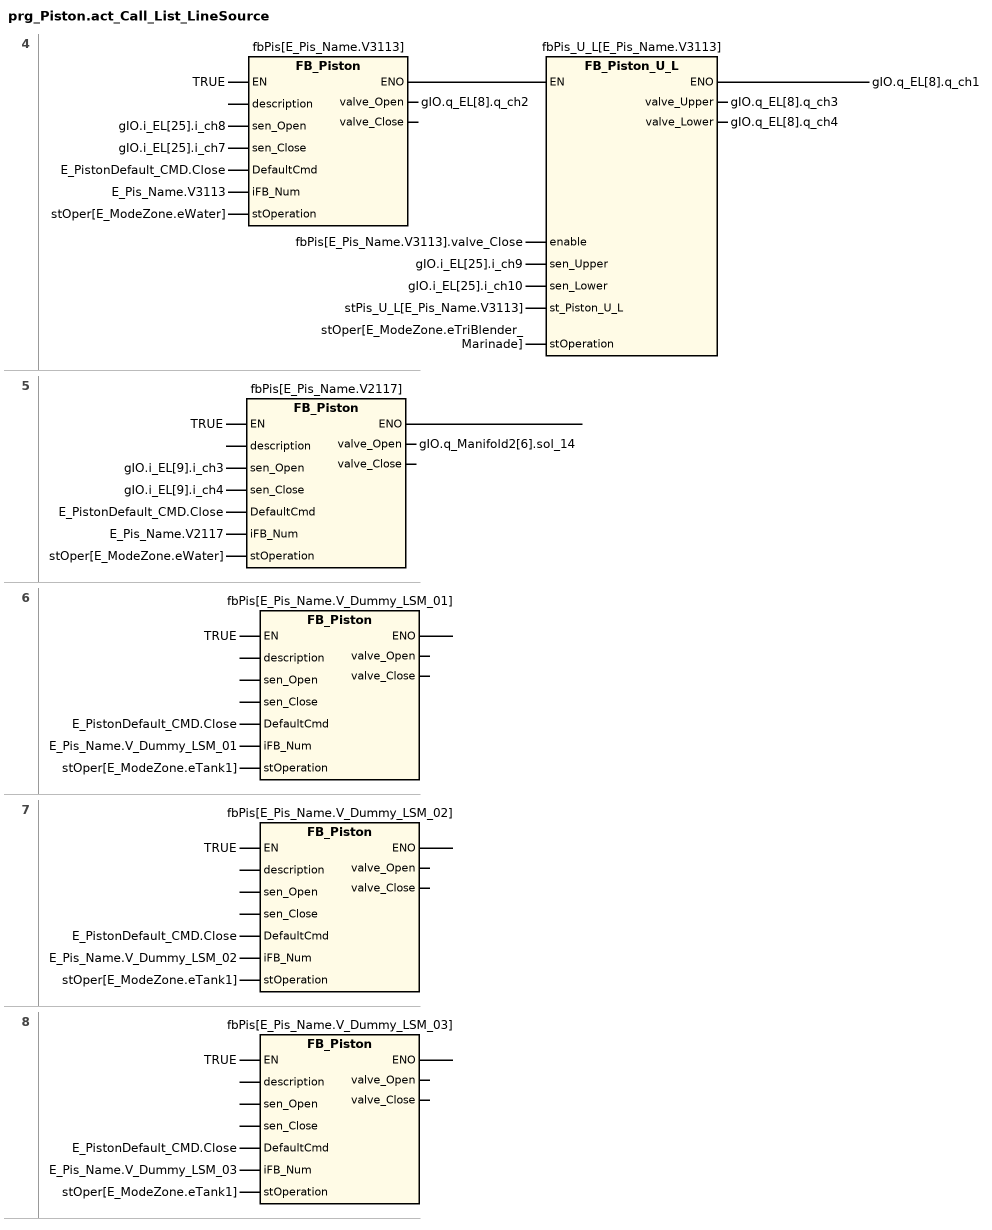
// NETWORK 4
fbPis[E_Pis_Name.V3113](
    sen_Open := gIO.i_EL[25].i_ch8,
    sen_Close := gIO.i_EL[25].i_ch7,
    DefaultCmd := E_PistonDefault_CMD.Close,
    iFB_Num := E_Pis_Name.V3113,
    stOperation := stOper[E_ModeZone.eWater],
    valve_Open => gIO.q_EL[8].q_ch2); // FB_Piston
fbPis_U_L[E_Pis_Name.V3113](
    enable := fbPis[E_Pis_Name.V3113].valve_Close,
    sen_Upper := gIO.i_EL[25].i_ch9,
    sen_Lower := gIO.i_EL[25].i_ch10,
    st_Piston_U_L := stPis_U_L[E_Pis_Name.V3113],
    stOperation := stOper[E_ModeZone.eTriBlender_Marinade],
    valve_Upper => gIO.q_EL[8].q_ch3,
    valve_Lower => gIO.q_EL[8].q_ch4); // FB_Piston_U_L
gIO.q_EL[8].q_ch1 := TRUE;

// NETWORK 5
fbPis[E_Pis_Name.V2117](
    sen_Open := gIO.i_EL[9].i_ch3,
    sen_Close := gIO.i_EL[9].i_ch4,
    DefaultCmd := E_PistonDefault_CMD.Close,
    iFB_Num := E_Pis_Name.V2117,
    stOperation := stOper[E_ModeZone.eWater],
    valve_Open => gIO.q_Manifold2[6].sol_14); // FB_Piston

// NETWORK 6
fbPis[E_Pis_Name.V_Dummy_LSM_01](
    DefaultCmd := E_PistonDefault_CMD.Close,
    iFB_Num := E_Pis_Name.V_Dummy_LSM_01,
    stOperation := stOper[E_ModeZone.eTank1]); // FB_Piston

// NETWORK 7
fbPis[E_Pis_Name.V_Dummy_LSM_02](
    DefaultCmd := E_PistonDefault_CMD.Close,
    iFB_Num := E_Pis_Name.V_Dummy_LSM_02,
    stOperation := stOper[E_ModeZone.eTank1]); // FB_Piston

// NETWORK 8
fbPis[E_Pis_Name.V_Dummy_LSM_03](
    DefaultCmd := E_PistonDefault_CMD.Close,
    iFB_Num := E_Pis_Name.V_Dummy_LSM_03,
    stOperation := stOper[E_ModeZone.eTank1]); // FB_Piston

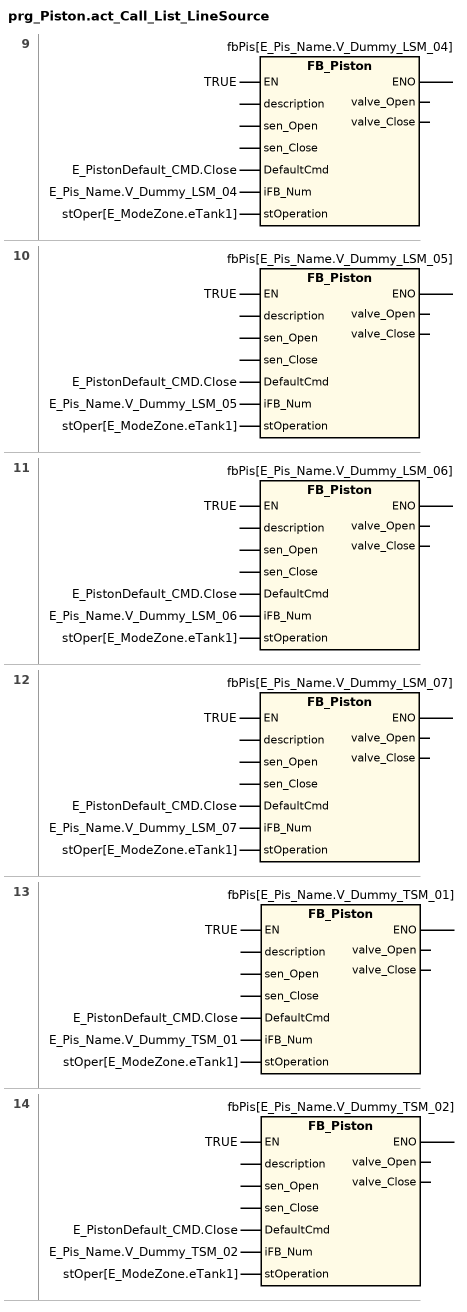
// NETWORK 9
fbPis[E_Pis_Name.V_Dummy_LSM_04](
    DefaultCmd := E_PistonDefault_CMD.Close,
    iFB_Num := E_Pis_Name.V_Dummy_LSM_04,
    stOperation := stOper[E_ModeZone.eTank1]); // FB_Piston

// NETWORK 10
fbPis[E_Pis_Name.V_Dummy_LSM_05](
    DefaultCmd := E_PistonDefault_CMD.Close,
    iFB_Num := E_Pis_Name.V_Dummy_LSM_05,
    stOperation := stOper[E_ModeZone.eTank1]); // FB_Piston

// NETWORK 11
fbPis[E_Pis_Name.V_Dummy_LSM_06](
    DefaultCmd := E_PistonDefault_CMD.Close,
    iFB_Num := E_Pis_Name.V_Dummy_LSM_06,
    stOperation := stOper[E_ModeZone.eTank1]); // FB_Piston

// NETWORK 12
fbPis[E_Pis_Name.V_Dummy_LSM_07](
    DefaultCmd := E_PistonDefault_CMD.Close,
    iFB_Num := E_Pis_Name.V_Dummy_LSM_07,
    stOperation := stOper[E_ModeZone.eTank1]); // FB_Piston

// NETWORK 13
fbPis[E_Pis_Name.V_Dummy_TSM_01](
    DefaultCmd := E_PistonDefault_CMD.Close,
    iFB_Num := E_Pis_Name.V_Dummy_TSM_01,
    stOperation := stOper[E_ModeZone.eTank1]); // FB_Piston

// NETWORK 14
fbPis[E_Pis_Name.V_Dummy_TSM_02](
    DefaultCmd := E_PistonDefault_CMD.Close,
    iFB_Num := E_Pis_Name.V_Dummy_TSM_02,
    stOperation := stOper[E_ModeZone.eTank1]); // FB_Piston

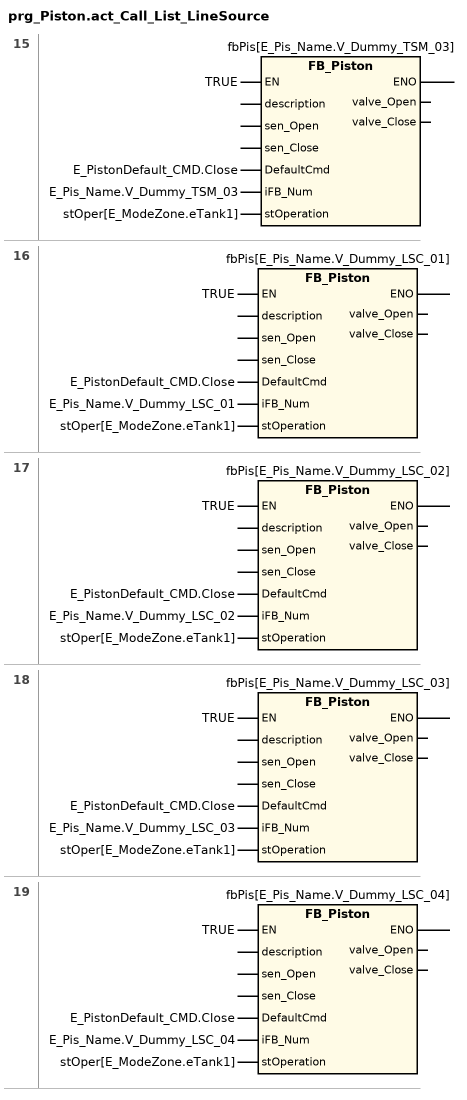
// NETWORK 15
fbPis[E_Pis_Name.V_Dummy_TSM_03](
    DefaultCmd := E_PistonDefault_CMD.Close,
    iFB_Num := E_Pis_Name.V_Dummy_TSM_03,
    stOperation := stOper[E_ModeZone.eTank1]); // FB_Piston

// NETWORK 16
fbPis[E_Pis_Name.V_Dummy_LSC_01](
    DefaultCmd := E_PistonDefault_CMD.Close,
    iFB_Num := E_Pis_Name.V_Dummy_LSC_01,
    stOperation := stOper[E_ModeZone.eTank1]); // FB_Piston

// NETWORK 17
fbPis[E_Pis_Name.V_Dummy_LSC_02](
    DefaultCmd := E_PistonDefault_CMD.Close,
    iFB_Num := E_Pis_Name.V_Dummy_LSC_02,
    stOperation := stOper[E_ModeZone.eTank1]); // FB_Piston

// NETWORK 18
fbPis[E_Pis_Name.V_Dummy_LSC_03](
    DefaultCmd := E_PistonDefault_CMD.Close,
    iFB_Num := E_Pis_Name.V_Dummy_LSC_03,
    stOperation := stOper[E_ModeZone.eTank1]); // FB_Piston

// NETWORK 19
fbPis[E_Pis_Name.V_Dummy_LSC_04](
    DefaultCmd := E_PistonDefault_CMD.Close,
    iFB_Num := E_Pis_Name.V_Dummy_LSC_04,
    stOperation := stOper[E_ModeZone.eTank1]); // FB_Piston
END_ACTION

ACTION act_Call_List_LineTarget:
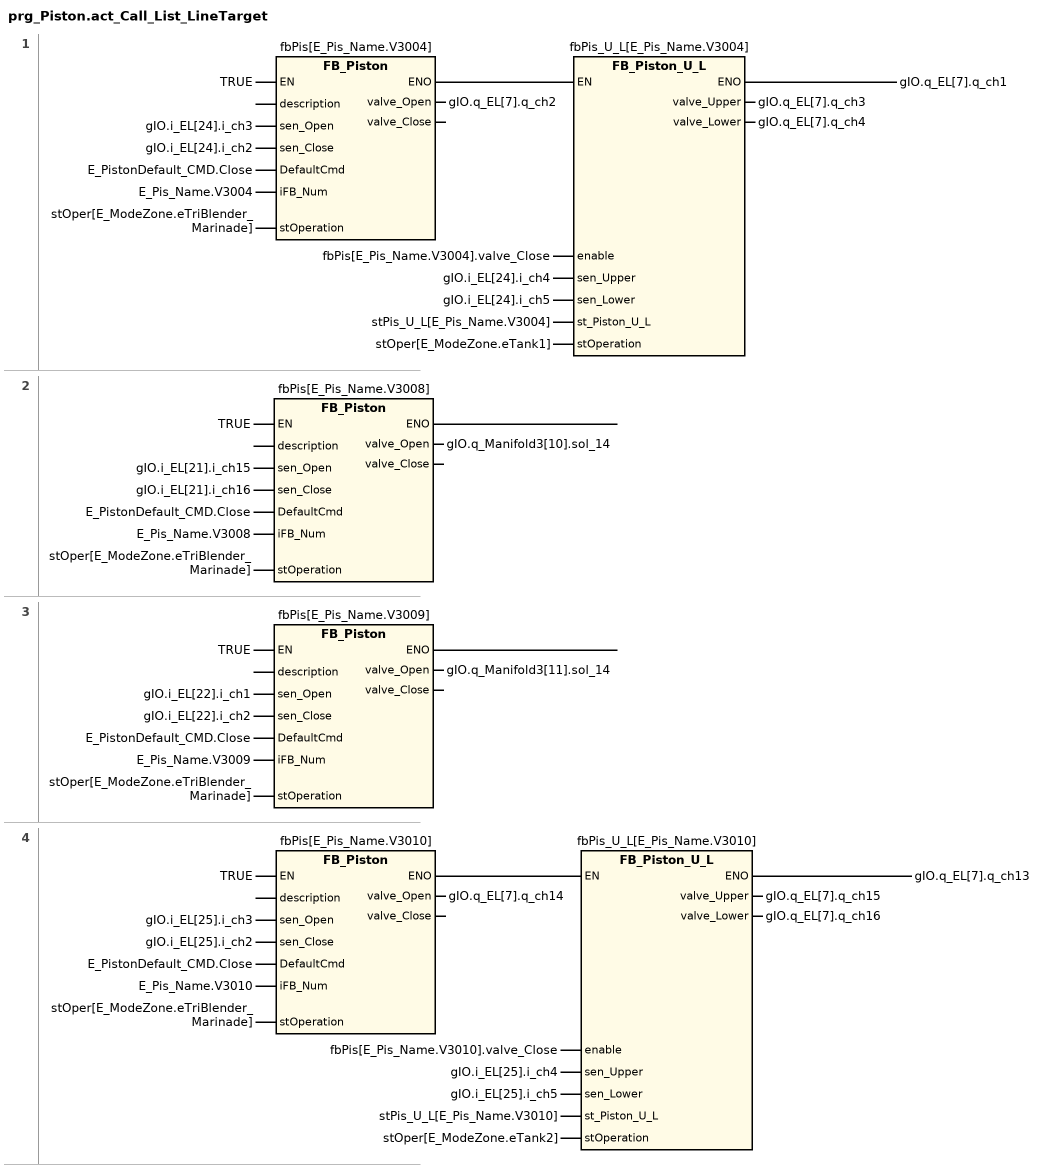
// NETWORK 1
fbPis[E_Pis_Name.V3004](
    sen_Open := gIO.i_EL[24].i_ch3,
    sen_Close := gIO.i_EL[24].i_ch2,
    DefaultCmd := E_PistonDefault_CMD.Close,
    iFB_Num := E_Pis_Name.V3004,
    stOperation := stOper[E_ModeZone.eTriBlender_Marinade],
    valve_Open => gIO.q_EL[7].q_ch2); // FB_Piston
fbPis_U_L[E_Pis_Name.V3004](
    enable := fbPis[E_Pis_Name.V3004].valve_Close,
    sen_Upper := gIO.i_EL[24].i_ch4,
    sen_Lower := gIO.i_EL[24].i_ch5,
    st_Piston_U_L := stPis_U_L[E_Pis_Name.V3004],
    stOperation := stOper[E_ModeZone.eTank1],
    valve_Upper => gIO.q_EL[7].q_ch3,
    valve_Lower => gIO.q_EL[7].q_ch4); // FB_Piston_U_L
gIO.q_EL[7].q_ch1 := TRUE;

// NETWORK 2
fbPis[E_Pis_Name.V3008](
    sen_Open := gIO.i_EL[21].i_ch15,
    sen_Close := gIO.i_EL[21].i_ch16,
    DefaultCmd := E_PistonDefault_CMD.Close,
    iFB_Num := E_Pis_Name.V3008,
    stOperation := stOper[E_ModeZone.eTriBlender_Marinade],
    valve_Open => gIO.q_Manifold3[10].sol_14); // FB_Piston

// NETWORK 3
fbPis[E_Pis_Name.V3009](
    sen_Open := gIO.i_EL[22].i_ch1,
    sen_Close := gIO.i_EL[22].i_ch2,
    DefaultCmd := E_PistonDefault_CMD.Close,
    iFB_Num := E_Pis_Name.V3009,
    stOperation := stOper[E_ModeZone.eTriBlender_Marinade],
    valve_Open => gIO.q_Manifold3[11].sol_14); // FB_Piston

// NETWORK 4
fbPis[E_Pis_Name.V3010](
    sen_Open := gIO.i_EL[25].i_ch3,
    sen_Close := gIO.i_EL[25].i_ch2,
    DefaultCmd := E_PistonDefault_CMD.Close,
    iFB_Num := E_Pis_Name.V3010,
    stOperation := stOper[E_ModeZone.eTriBlender_Marinade],
    valve_Open => gIO.q_EL[7].q_ch14); // FB_Piston
fbPis_U_L[E_Pis_Name.V3010](
    enable := fbPis[E_Pis_Name.V3010].valve_Close,
    sen_Upper := gIO.i_EL[25].i_ch4,
    sen_Lower := gIO.i_EL[25].i_ch5,
    st_Piston_U_L := stPis_U_L[E_Pis_Name.V3010],
    stOperation := stOper[E_ModeZone.eTank2],
    valve_Upper => gIO.q_EL[7].q_ch15,
    valve_Lower => gIO.q_EL[7].q_ch16); // FB_Piston_U_L
gIO.q_EL[7].q_ch13 := TRUE;

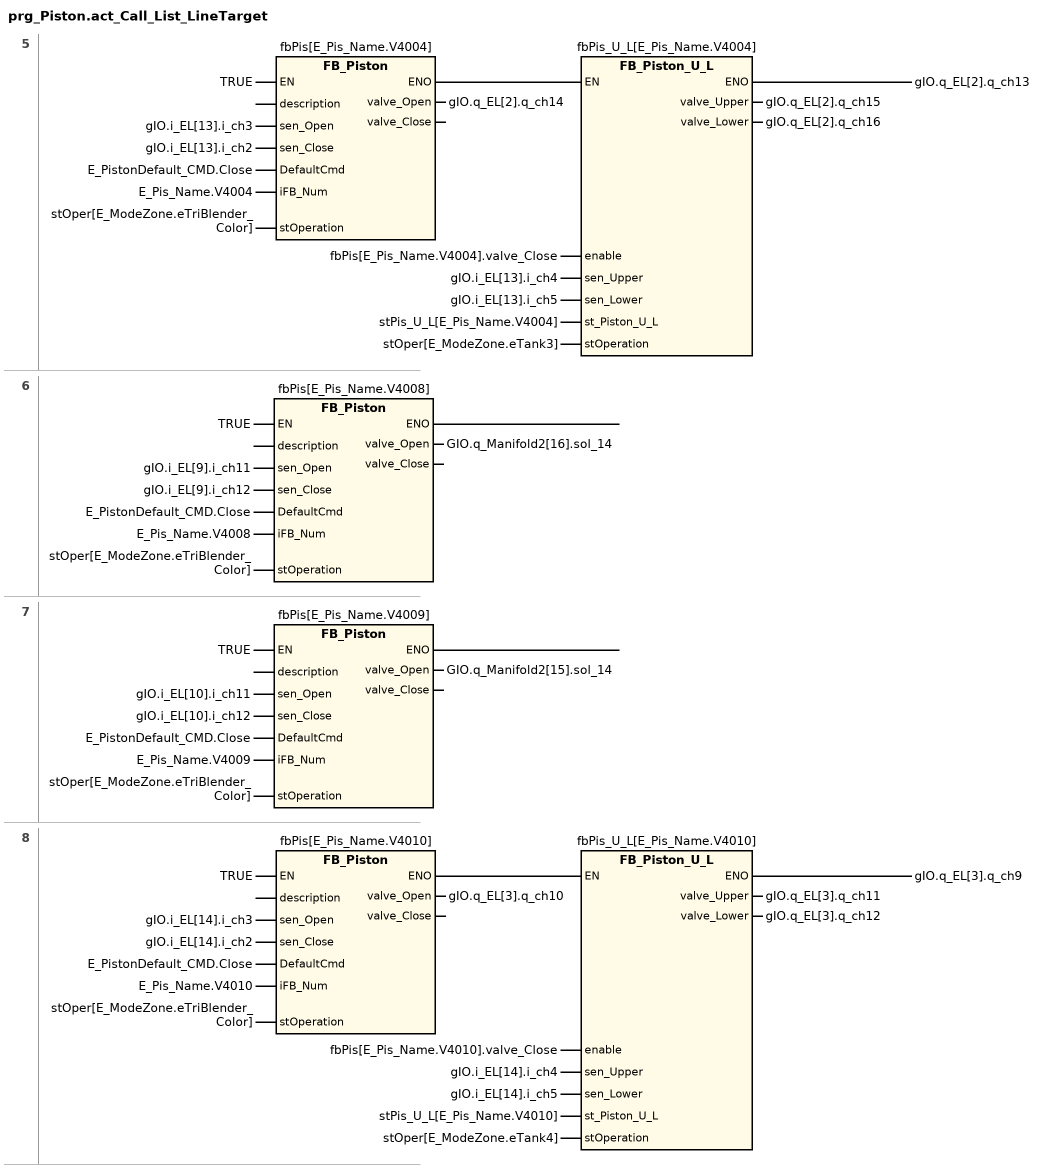
// NETWORK 5
fbPis[E_Pis_Name.V4004](
    sen_Open := gIO.i_EL[13].i_ch3,
    sen_Close := gIO.i_EL[13].i_ch2,
    DefaultCmd := E_PistonDefault_CMD.Close,
    iFB_Num := E_Pis_Name.V4004,
    stOperation := stOper[E_ModeZone.eTriBlender_Color],
    valve_Open => gIO.q_EL[2].q_ch14); // FB_Piston
fbPis_U_L[E_Pis_Name.V4004](
    enable := fbPis[E_Pis_Name.V4004].valve_Close,
    sen_Upper := gIO.i_EL[13].i_ch4,
    sen_Lower := gIO.i_EL[13].i_ch5,
    st_Piston_U_L := stPis_U_L[E_Pis_Name.V4004],
    stOperation := stOper[E_ModeZone.eTank3],
    valve_Upper => gIO.q_EL[2].q_ch15,
    valve_Lower => gIO.q_EL[2].q_ch16); // FB_Piston_U_L
gIO.q_EL[2].q_ch13 := TRUE;

// NETWORK 6
fbPis[E_Pis_Name.V4008](
    sen_Open := gIO.i_EL[9].i_ch11,
    sen_Close := gIO.i_EL[9].i_ch12,
    DefaultCmd := E_PistonDefault_CMD.Close,
    iFB_Num := E_Pis_Name.V4008,
    stOperation := stOper[E_ModeZone.eTriBlender_Color],
    valve_Open => GIO.q_Manifold2[16].sol_14); // FB_Piston

// NETWORK 7
fbPis[E_Pis_Name.V4009](
    sen_Open := gIO.i_EL[10].i_ch11,
    sen_Close := gIO.i_EL[10].i_ch12,
    DefaultCmd := E_PistonDefault_CMD.Close,
    iFB_Num := E_Pis_Name.V4009,
    stOperation := stOper[E_ModeZone.eTriBlender_Color],
    valve_Open => GIO.q_Manifold2[15].sol_14); // FB_Piston

// NETWORK 8
fbPis[E_Pis_Name.V4010](
    sen_Open := gIO.i_EL[14].i_ch3,
    sen_Close := gIO.i_EL[14].i_ch2,
    DefaultCmd := E_PistonDefault_CMD.Close,
    iFB_Num := E_Pis_Name.V4010,
    stOperation := stOper[E_ModeZone.eTriBlender_Color],
    valve_Open => gIO.q_EL[3].q_ch10); // FB_Piston
fbPis_U_L[E_Pis_Name.V4010](
    enable := fbPis[E_Pis_Name.V4010].valve_Close,
    sen_Upper := gIO.i_EL[14].i_ch4,
    sen_Lower := gIO.i_EL[14].i_ch5,
    st_Piston_U_L := stPis_U_L[E_Pis_Name.V4010],
    stOperation := stOper[E_ModeZone.eTank4],
    valve_Upper => gIO.q_EL[3].q_ch11,
    valve_Lower => gIO.q_EL[3].q_ch12); // FB_Piston_U_L
gIO.q_EL[3].q_ch9 := TRUE;

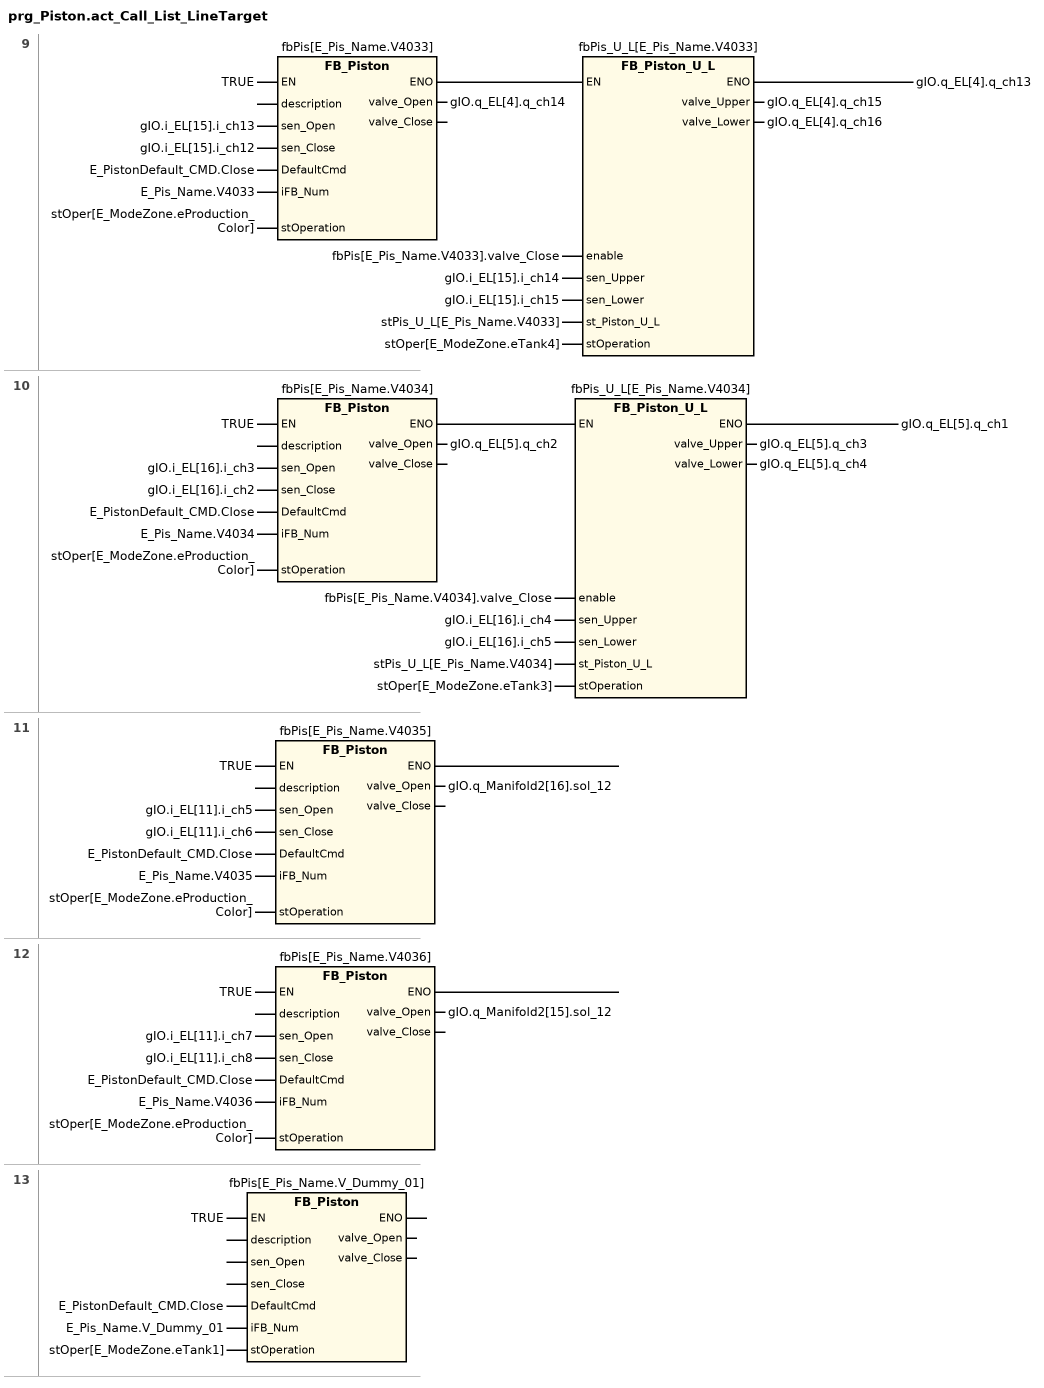
// NETWORK 9
fbPis[E_Pis_Name.V4033](
    sen_Open := gIO.i_EL[15].i_ch13,
    sen_Close := gIO.i_EL[15].i_ch12,
    DefaultCmd := E_PistonDefault_CMD.Close,
    iFB_Num := E_Pis_Name.V4033,
    stOperation := stOper[E_ModeZone.eProduction_Color],
    valve_Open => gIO.q_EL[4].q_ch14); // FB_Piston
fbPis_U_L[E_Pis_Name.V4033](
    enable := fbPis[E_Pis_Name.V4033].valve_Close,
    sen_Upper := gIO.i_EL[15].i_ch14,
    sen_Lower := gIO.i_EL[15].i_ch15,
    st_Piston_U_L := stPis_U_L[E_Pis_Name.V4033],
    stOperation := stOper[E_ModeZone.eTank4],
    valve_Upper => gIO.q_EL[4].q_ch15,
    valve_Lower => gIO.q_EL[4].q_ch16); // FB_Piston_U_L
gIO.q_EL[4].q_ch13 := TRUE;

// NETWORK 10
fbPis[E_Pis_Name.V4034](
    sen_Open := gIO.i_EL[16].i_ch3,
    sen_Close := gIO.i_EL[16].i_ch2,
    DefaultCmd := E_PistonDefault_CMD.Close,
    iFB_Num := E_Pis_Name.V4034,
    stOperation := stOper[E_ModeZone.eProduction_Color],
    valve_Open => gIO.q_EL[5].q_ch2); // FB_Piston
fbPis_U_L[E_Pis_Name.V4034](
    enable := fbPis[E_Pis_Name.V4034].valve_Close,
    sen_Upper := gIO.i_EL[16].i_ch4,
    sen_Lower := gIO.i_EL[16].i_ch5,
    st_Piston_U_L := stPis_U_L[E_Pis_Name.V4034],
    stOperation := stOper[E_ModeZone.eTank3],
    valve_Upper => gIO.q_EL[5].q_ch3,
    valve_Lower => gIO.q_EL[5].q_ch4); // FB_Piston_U_L
gIO.q_EL[5].q_ch1 := TRUE;

// NETWORK 11
fbPis[E_Pis_Name.V4035](
    sen_Open := gIO.i_EL[11].i_ch5,
    sen_Close := gIO.i_EL[11].i_ch6,
    DefaultCmd := E_PistonDefault_CMD.Close,
    iFB_Num := E_Pis_Name.V4035,
    stOperation := stOper[E_ModeZone.eProduction_Color],
    valve_Open => gIO.q_Manifold2[16].sol_12); // FB_Piston

// NETWORK 12
fbPis[E_Pis_Name.V4036](
    sen_Open := gIO.i_EL[11].i_ch7,
    sen_Close := gIO.i_EL[11].i_ch8,
    DefaultCmd := E_PistonDefault_CMD.Close,
    iFB_Num := E_Pis_Name.V4036,
    stOperation := stOper[E_ModeZone.eProduction_Color],
    valve_Open => gIO.q_Manifold2[15].sol_12); // FB_Piston

// NETWORK 13
fbPis[E_Pis_Name.V_Dummy_01](
    DefaultCmd := E_PistonDefault_CMD.Close,
    iFB_Num := E_Pis_Name.V_Dummy_01,
    stOperation := stOper[E_ModeZone.eTank1]); // FB_Piston

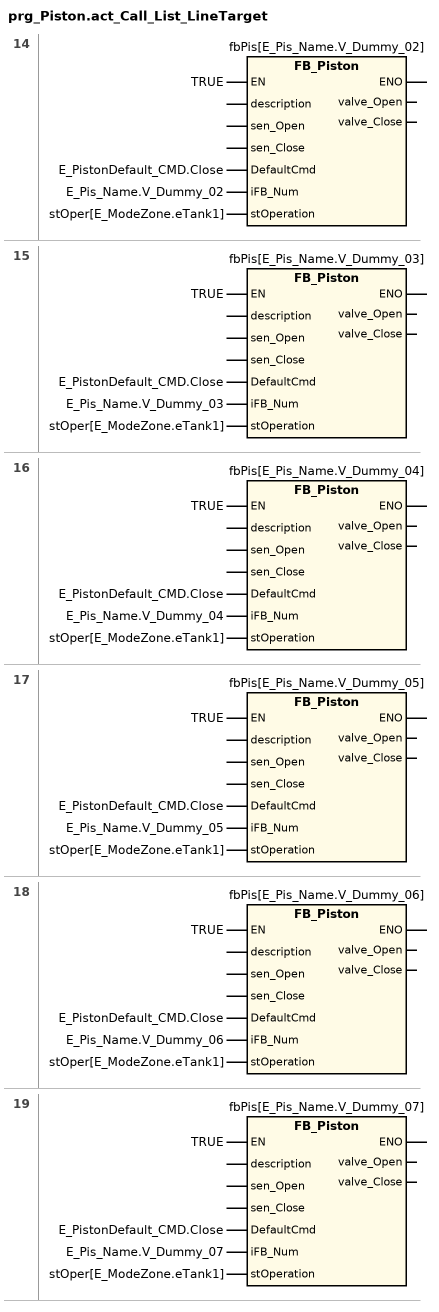
// NETWORK 14
fbPis[E_Pis_Name.V_Dummy_02](
    DefaultCmd := E_PistonDefault_CMD.Close,
    iFB_Num := E_Pis_Name.V_Dummy_02,
    stOperation := stOper[E_ModeZone.eTank1]); // FB_Piston

// NETWORK 15
fbPis[E_Pis_Name.V_Dummy_03](
    DefaultCmd := E_PistonDefault_CMD.Close,
    iFB_Num := E_Pis_Name.V_Dummy_03,
    stOperation := stOper[E_ModeZone.eTank1]); // FB_Piston

// NETWORK 16
fbPis[E_Pis_Name.V_Dummy_04](
    DefaultCmd := E_PistonDefault_CMD.Close,
    iFB_Num := E_Pis_Name.V_Dummy_04,
    stOperation := stOper[E_ModeZone.eTank1]); // FB_Piston

// NETWORK 17
fbPis[E_Pis_Name.V_Dummy_05](
    DefaultCmd := E_PistonDefault_CMD.Close,
    iFB_Num := E_Pis_Name.V_Dummy_05,
    stOperation := stOper[E_ModeZone.eTank1]); // FB_Piston

// NETWORK 18
fbPis[E_Pis_Name.V_Dummy_06](
    DefaultCmd := E_PistonDefault_CMD.Close,
    iFB_Num := E_Pis_Name.V_Dummy_06,
    stOperation := stOper[E_ModeZone.eTank1]); // FB_Piston

// NETWORK 19
fbPis[E_Pis_Name.V_Dummy_07](
    DefaultCmd := E_PistonDefault_CMD.Close,
    iFB_Num := E_Pis_Name.V_Dummy_07,
    stOperation := stOper[E_ModeZone.eTank1]); // FB_Piston

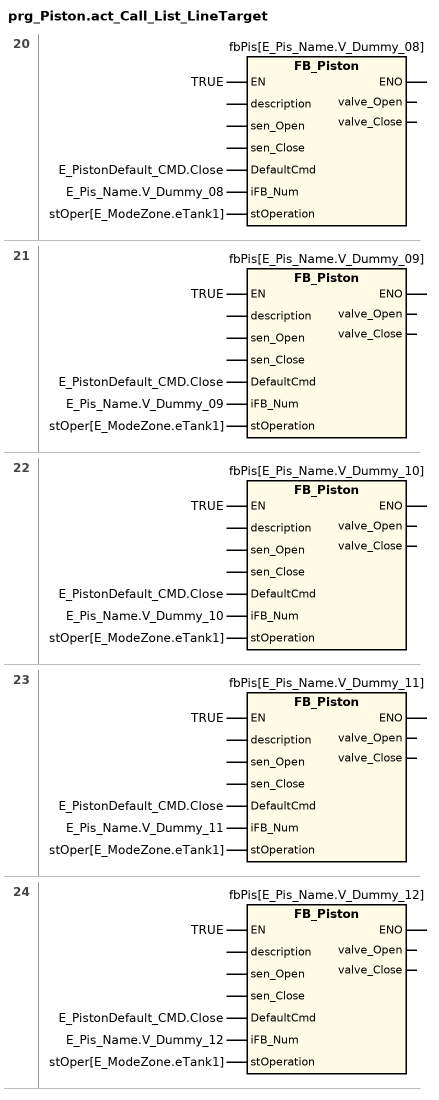
// NETWORK 20
fbPis[E_Pis_Name.V_Dummy_08](
    DefaultCmd := E_PistonDefault_CMD.Close,
    iFB_Num := E_Pis_Name.V_Dummy_08,
    stOperation := stOper[E_ModeZone.eTank1]); // FB_Piston

// NETWORK 21
fbPis[E_Pis_Name.V_Dummy_09](
    DefaultCmd := E_PistonDefault_CMD.Close,
    iFB_Num := E_Pis_Name.V_Dummy_09,
    stOperation := stOper[E_ModeZone.eTank1]); // FB_Piston

// NETWORK 22
fbPis[E_Pis_Name.V_Dummy_10](
    DefaultCmd := E_PistonDefault_CMD.Close,
    iFB_Num := E_Pis_Name.V_Dummy_10,
    stOperation := stOper[E_ModeZone.eTank1]); // FB_Piston

// NETWORK 23
fbPis[E_Pis_Name.V_Dummy_11](
    DefaultCmd := E_PistonDefault_CMD.Close,
    iFB_Num := E_Pis_Name.V_Dummy_11,
    stOperation := stOper[E_ModeZone.eTank1]); // FB_Piston

// NETWORK 24
fbPis[E_Pis_Name.V_Dummy_12](
    DefaultCmd := E_PistonDefault_CMD.Close,
    iFB_Num := E_Pis_Name.V_Dummy_12,
    stOperation := stOper[E_ModeZone.eTank1]); // FB_Piston
END_ACTION

ACTION act_Call_list_TanksColor:
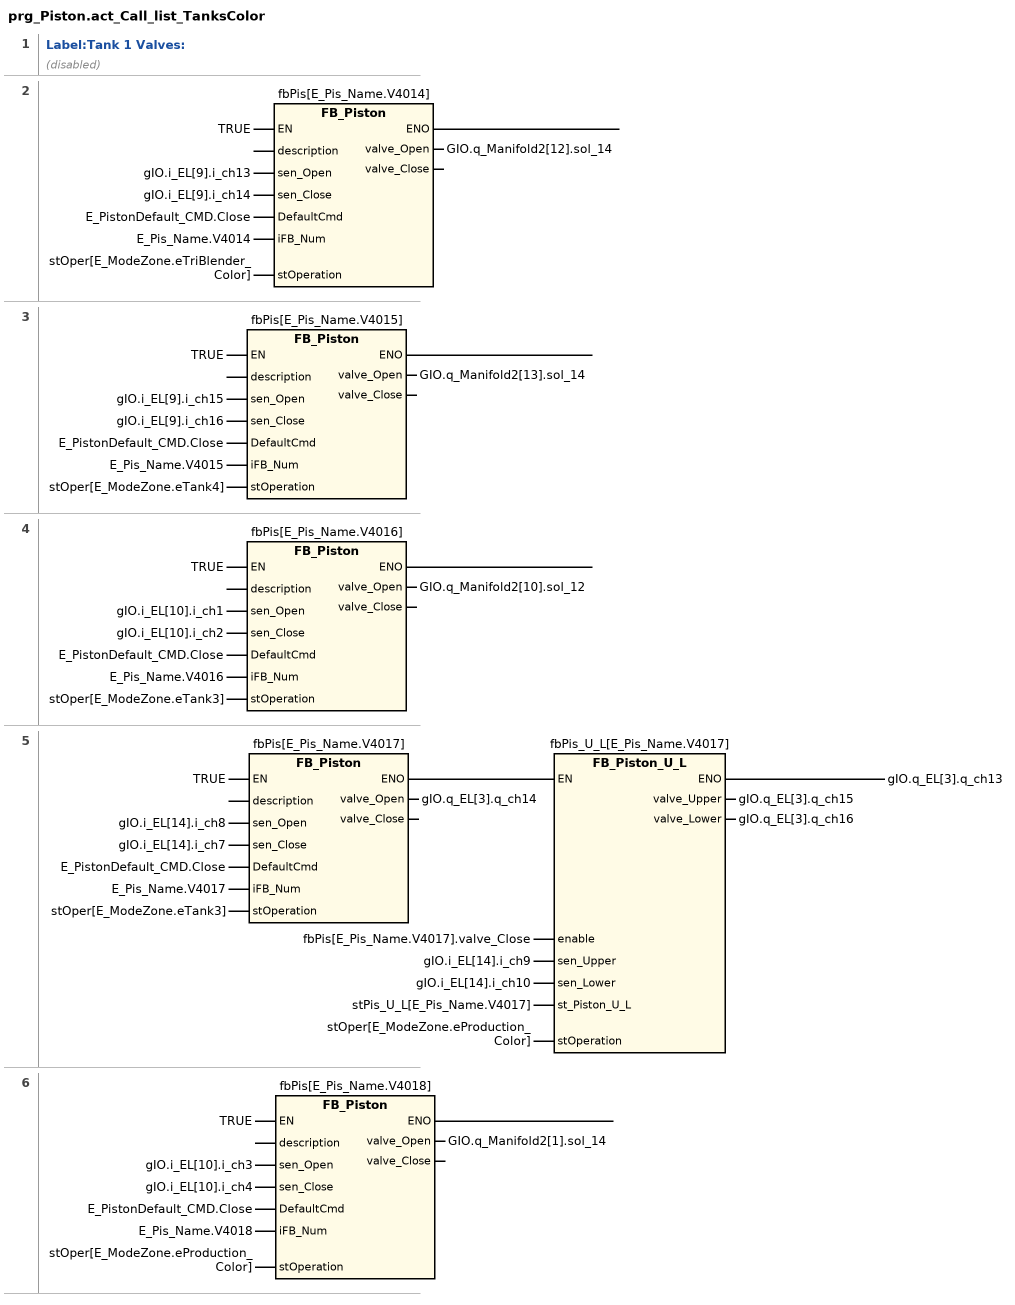
// NETWORK 1 (disabled)
// label: Label:Tank 1 Valves

// NETWORK 2
fbPis[E_Pis_Name.V4014](
    sen_Open := gIO.i_EL[9].i_ch13,
    sen_Close := gIO.i_EL[9].i_ch14,
    DefaultCmd := E_PistonDefault_CMD.Close,
    iFB_Num := E_Pis_Name.V4014,
    stOperation := stOper[E_ModeZone.eTriBlender_Color],
    valve_Open => GIO.q_Manifold2[12].sol_14); // FB_Piston

// NETWORK 3
fbPis[E_Pis_Name.V4015](
    sen_Open := gIO.i_EL[9].i_ch15,
    sen_Close := gIO.i_EL[9].i_ch16,
    DefaultCmd := E_PistonDefault_CMD.Close,
    iFB_Num := E_Pis_Name.V4015,
    stOperation := stOper[E_ModeZone.eTank4],
    valve_Open => GIO.q_Manifold2[13].sol_14); // FB_Piston

// NETWORK 4
fbPis[E_Pis_Name.V4016](
    sen_Open := gIO.i_EL[10].i_ch1,
    sen_Close := gIO.i_EL[10].i_ch2,
    DefaultCmd := E_PistonDefault_CMD.Close,
    iFB_Num := E_Pis_Name.V4016,
    stOperation := stOper[E_ModeZone.eTank3],
    valve_Open => GIO.q_Manifold2[10].sol_12); // FB_Piston

// NETWORK 5
fbPis[E_Pis_Name.V4017](
    sen_Open := gIO.i_EL[14].i_ch8,
    sen_Close := gIO.i_EL[14].i_ch7,
    DefaultCmd := E_PistonDefault_CMD.Close,
    iFB_Num := E_Pis_Name.V4017,
    stOperation := stOper[E_ModeZone.eTank3],
    valve_Open => gIO.q_EL[3].q_ch14); // FB_Piston
fbPis_U_L[E_Pis_Name.V4017](
    enable := fbPis[E_Pis_Name.V4017].valve_Close,
    sen_Upper := gIO.i_EL[14].i_ch9,
    sen_Lower := gIO.i_EL[14].i_ch10,
    st_Piston_U_L := stPis_U_L[E_Pis_Name.V4017],
    stOperation := stOper[E_ModeZone.eProduction_Color],
    valve_Upper => gIO.q_EL[3].q_ch15,
    valve_Lower => gIO.q_EL[3].q_ch16); // FB_Piston_U_L
gIO.q_EL[3].q_ch13 := TRUE;

// NETWORK 6
fbPis[E_Pis_Name.V4018](
    sen_Open := gIO.i_EL[10].i_ch3,
    sen_Close := gIO.i_EL[10].i_ch4,
    DefaultCmd := E_PistonDefault_CMD.Close,
    iFB_Num := E_Pis_Name.V4018,
    stOperation := stOper[E_ModeZone.eProduction_Color],
    valve_Open => GIO.q_Manifold2[1].sol_14); // FB_Piston

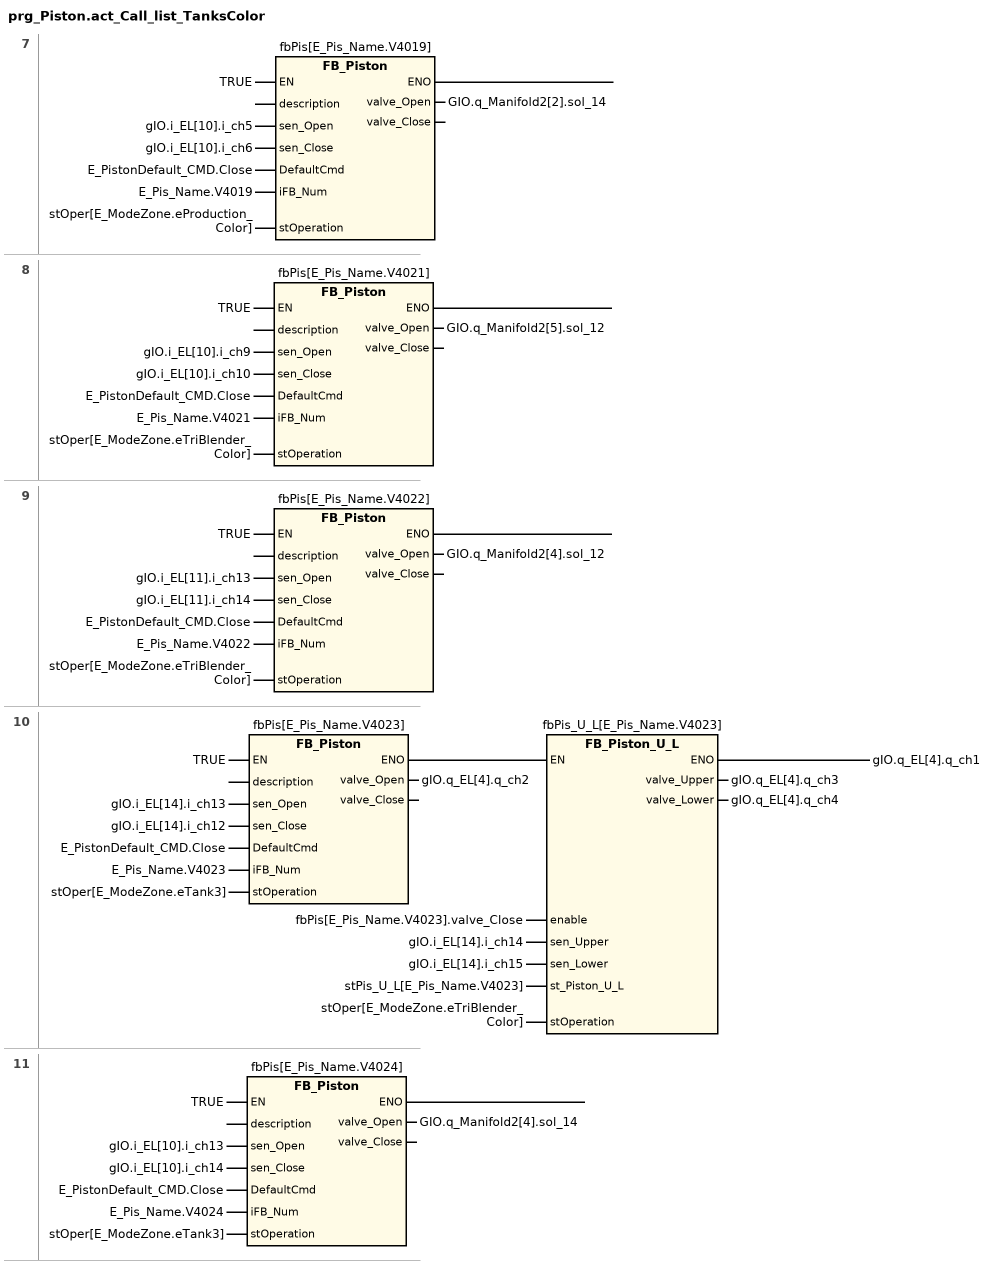
// NETWORK 7
fbPis[E_Pis_Name.V4019](
    sen_Open := gIO.i_EL[10].i_ch5,
    sen_Close := gIO.i_EL[10].i_ch6,
    DefaultCmd := E_PistonDefault_CMD.Close,
    iFB_Num := E_Pis_Name.V4019,
    stOperation := stOper[E_ModeZone.eProduction_Color],
    valve_Open => GIO.q_Manifold2[2].sol_14); // FB_Piston

// NETWORK 8
fbPis[E_Pis_Name.V4021](
    sen_Open := gIO.i_EL[10].i_ch9,
    sen_Close := gIO.i_EL[10].i_ch10,
    DefaultCmd := E_PistonDefault_CMD.Close,
    iFB_Num := E_Pis_Name.V4021,
    stOperation := stOper[E_ModeZone.eTriBlender_Color],
    valve_Open => GIO.q_Manifold2[5].sol_12); // FB_Piston

// NETWORK 9
fbPis[E_Pis_Name.V4022](
    sen_Open := gIO.i_EL[11].i_ch13,
    sen_Close := gIO.i_EL[11].i_ch14,
    DefaultCmd := E_PistonDefault_CMD.Close,
    iFB_Num := E_Pis_Name.V4022,
    stOperation := stOper[E_ModeZone.eTriBlender_Color],
    valve_Open => GIO.q_Manifold2[4].sol_12); // FB_Piston

// NETWORK 10
fbPis[E_Pis_Name.V4023](
    sen_Open := gIO.i_EL[14].i_ch13,
    sen_Close := gIO.i_EL[14].i_ch12,
    DefaultCmd := E_PistonDefault_CMD.Close,
    iFB_Num := E_Pis_Name.V4023,
    stOperation := stOper[E_ModeZone.eTank3],
    valve_Open => gIO.q_EL[4].q_ch2); // FB_Piston
fbPis_U_L[E_Pis_Name.V4023](
    enable := fbPis[E_Pis_Name.V4023].valve_Close,
    sen_Upper := gIO.i_EL[14].i_ch14,
    sen_Lower := gIO.i_EL[14].i_ch15,
    st_Piston_U_L := stPis_U_L[E_Pis_Name.V4023],
    stOperation := stOper[E_ModeZone.eTriBlender_Color],
    valve_Upper => gIO.q_EL[4].q_ch3,
    valve_Lower => gIO.q_EL[4].q_ch4); // FB_Piston_U_L
gIO.q_EL[4].q_ch1 := TRUE;

// NETWORK 11
fbPis[E_Pis_Name.V4024](
    sen_Open := gIO.i_EL[10].i_ch13,
    sen_Close := gIO.i_EL[10].i_ch14,
    DefaultCmd := E_PistonDefault_CMD.Close,
    iFB_Num := E_Pis_Name.V4024,
    stOperation := stOper[E_ModeZone.eTank3],
    valve_Open => GIO.q_Manifold2[4].sol_14); // FB_Piston

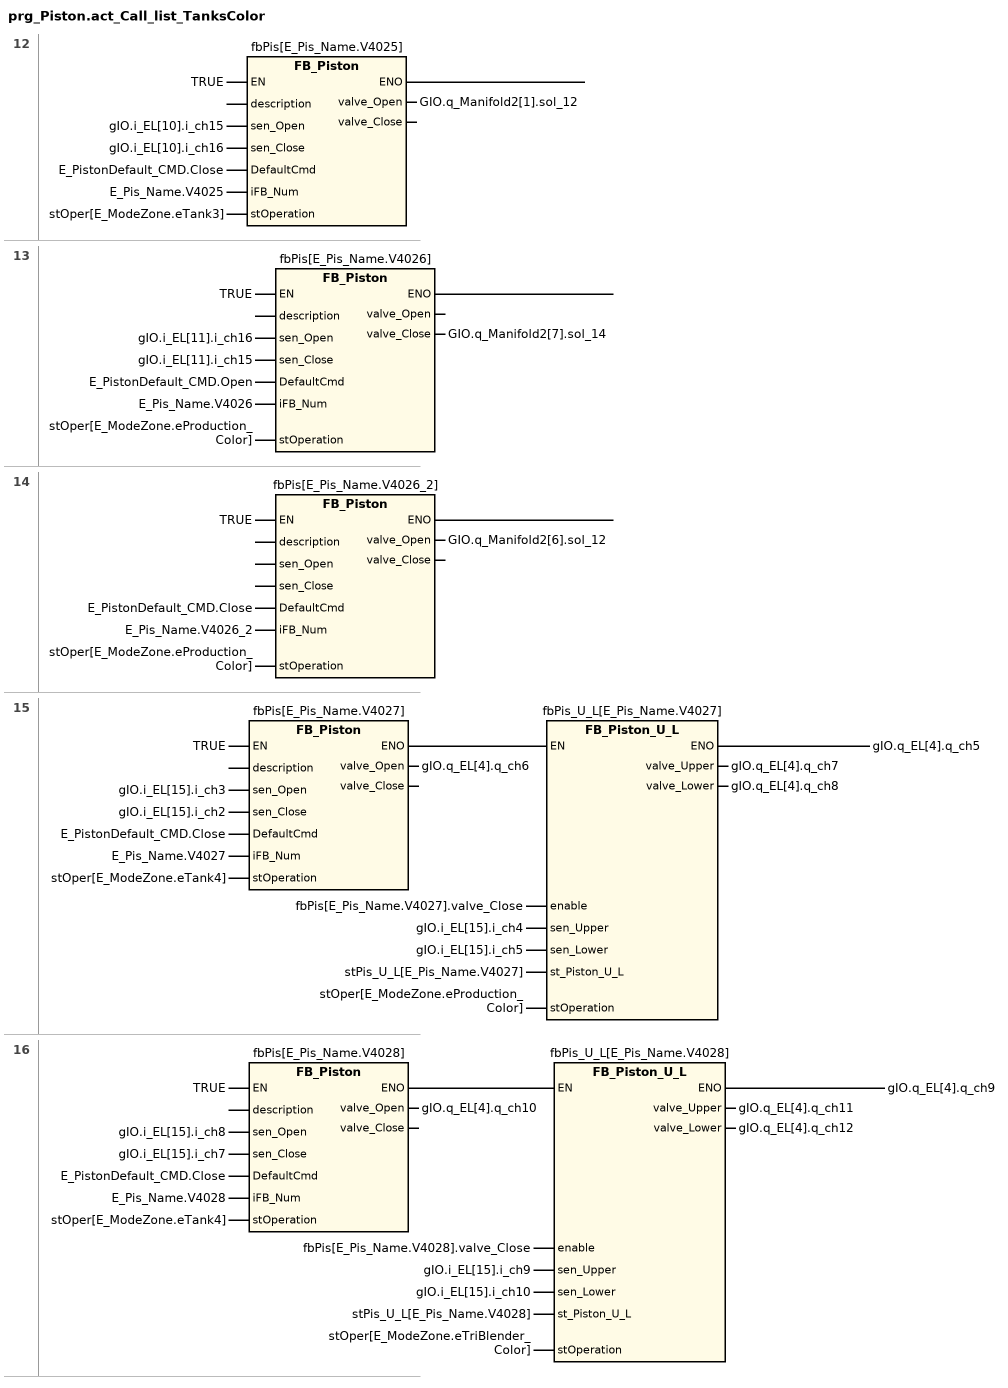
// NETWORK 12
fbPis[E_Pis_Name.V4025](
    sen_Open := gIO.i_EL[10].i_ch15,
    sen_Close := gIO.i_EL[10].i_ch16,
    DefaultCmd := E_PistonDefault_CMD.Close,
    iFB_Num := E_Pis_Name.V4025,
    stOperation := stOper[E_ModeZone.eTank3],
    valve_Open => GIO.q_Manifold2[1].sol_12); // FB_Piston

// NETWORK 13
fbPis[E_Pis_Name.V4026](
    sen_Open := gIO.i_EL[11].i_ch16,
    sen_Close := gIO.i_EL[11].i_ch15,
    DefaultCmd := E_PistonDefault_CMD.Open,
    iFB_Num := E_Pis_Name.V4026,
    stOperation := stOper[E_ModeZone.eProduction_Color],
    valve_Close => GIO.q_Manifold2[7].sol_14); // FB_Piston

// NETWORK 14
fbPis[E_Pis_Name.V4026_2](
    DefaultCmd := E_PistonDefault_CMD.Close,
    iFB_Num := E_Pis_Name.V4026_2,
    stOperation := stOper[E_ModeZone.eProduction_Color],
    valve_Open => GIO.q_Manifold2[6].sol_12); // FB_Piston

// NETWORK 15
fbPis[E_Pis_Name.V4027](
    sen_Open := gIO.i_EL[15].i_ch3,
    sen_Close := gIO.i_EL[15].i_ch2,
    DefaultCmd := E_PistonDefault_CMD.Close,
    iFB_Num := E_Pis_Name.V4027,
    stOperation := stOper[E_ModeZone.eTank4],
    valve_Open => gIO.q_EL[4].q_ch6); // FB_Piston
fbPis_U_L[E_Pis_Name.V4027](
    enable := fbPis[E_Pis_Name.V4027].valve_Close,
    sen_Upper := gIO.i_EL[15].i_ch4,
    sen_Lower := gIO.i_EL[15].i_ch5,
    st_Piston_U_L := stPis_U_L[E_Pis_Name.V4027],
    stOperation := stOper[E_ModeZone.eProduction_Color],
    valve_Upper => gIO.q_EL[4].q_ch7,
    valve_Lower => gIO.q_EL[4].q_ch8); // FB_Piston_U_L
gIO.q_EL[4].q_ch5 := TRUE;

// NETWORK 16
fbPis[E_Pis_Name.V4028](
    sen_Open := gIO.i_EL[15].i_ch8,
    sen_Close := gIO.i_EL[15].i_ch7,
    DefaultCmd := E_PistonDefault_CMD.Close,
    iFB_Num := E_Pis_Name.V4028,
    stOperation := stOper[E_ModeZone.eTank4],
    valve_Open => gIO.q_EL[4].q_ch10); // FB_Piston
fbPis_U_L[E_Pis_Name.V4028](
    enable := fbPis[E_Pis_Name.V4028].valve_Close,
    sen_Upper := gIO.i_EL[15].i_ch9,
    sen_Lower := gIO.i_EL[15].i_ch10,
    st_Piston_U_L := stPis_U_L[E_Pis_Name.V4028],
    stOperation := stOper[E_ModeZone.eTriBlender_Color],
    valve_Upper => gIO.q_EL[4].q_ch11,
    valve_Lower => gIO.q_EL[4].q_ch12); // FB_Piston_U_L
gIO.q_EL[4].q_ch9 := TRUE;

